{region 'Documentation'}
(*!
<summary>Reads a captured finding; the caller bounds the index by 8 subjects.</summary>
*)
{endregion}
METHOD PRIVATE IsFindingValid : BOOL //! TRUE when the selected captured finding satisfies the scenario metadata and diagnostic checks.
VAR_INPUT
    Index : UINT; //! One-based index in the retained isolated event capture.
    ExpectedName : STRING(GVL_Constants.NameLength); //! Independently authored Assertion name expected in the selected finding.
    ExpectedResult : E_Result; //! Independently authored finding result.
END_VAR
IsFindingValid := (FEvents[Index].SequenceId = UINT_TO_UDINT(Index))
    AND (FEvents[Index].Name = ExpectedName)
    AND (FEvents[Index].OwnerScope = E_OwnerScope.Assertion)
    AND (FEvents[Index].EventType = E_EventType.Result)
    AND (FEvents[Index].State = E_State.Running)
    AND (FEvents[Index].Result = ExpectedResult)
    AND (FEvents[Index].Message <> '');
END_METHOD

{region 'Documentation'}
(*!
<summary>Completes abort without asynchronous resources.</summary>
*)
{endregion}
METHOD PROTECTED ProcessAbort
VAR_INPUT
    Enable : BOOL; //! Phase permission supplied by the owning Test Case; FALSE does not authorize progression, while observation may continue.
END_VAR
IF Enable THEN
    CompleteAbort();
END_IF;
END_METHOD

{region 'Documentation'}
(*!
<summary>Latches checked observations before the next script step may proceed.</summary>
*)
{endregion}
METHOD PROTECTED ProcessAssertions
VAR_INPUT
    Enable : BOOL; //! Phase permission supplied by the owning Test Case; FALSE does not authorize progression, while observation may continue.
END_VAR
VAR
    Evaluate : BOOL;
END_VAR
Evaluate := Enable AND FObservationReady;
FEqualResult(Enable := Evaluate,
    State := State,
    IN := FEqualResultMatches);
FNotEqualResult(Enable := Evaluate,
    State := State,
    IN := FNotEqualResultMatches);
FLessThanResult(Enable := Evaluate,
    State := State,
    IN := FLessThanResultMatches);
FLessEqualResult(Enable := Evaluate,
    State := State,
    IN := FLessEqualResultMatches);
FGreaterThanResult(Enable := Evaluate,
    State := State,
    IN := FGreaterThanResultMatches);
FGreaterEqualResult(Enable := Evaluate,
    State := State,
    IN := FGreaterEqualResultMatches);
FInRangeResult(Enable := Evaluate,
    State := State,
    IN := FInRangeResultMatches);
FNotInRangeResult(Enable := Evaluate,
    State := State,
    IN := FNotInRangeResultMatches);
FCaptureIntegrity(Enable := Evaluate,
    State := State,
    IN := FCaptureIntegrityMatches);
FFindingDetails(Enable := Evaluate,
    State := State,
    IN := FFindingDetailsMatch);
IF Evaluate THEN
    FChecked := TRUE;
END_IF;
END_METHOD

{region 'Documentation'}
(*!
<summary>No Preparation phase is required.</summary>
*)
{endregion}
METHOD PROTECTED ProcessPreparations
VAR_INPUT
    // SA0033: Required hook; this test has no Preparation phase.
    {attribute 'analysis' := '-33'}
    Enable : BOOL; //! Phase permission supplied by the owning Test Case; FALSE does not authorize progression, while observation may continue.
END_VAR
END_METHOD

{region 'Documentation'}
(*!
<summary>Restarts the script and resets the checking Assertions.</summary>
*)
{endregion}
METHOD PROTECTED ProcessReset
FRow := EqualAtLowerBound;
FRowPrepared := FALSE;
FChecked := FALSE;
FObservationReady := FALSE;
FEqualResult.Reset();
FEqualResultMatches := TRUE;
FNotEqualResult.Reset();
FNotEqualResultMatches := TRUE;
FLessThanResult.Reset();
FLessThanResultMatches := TRUE;
FLessEqualResult.Reset();
FLessEqualResultMatches := TRUE;
FGreaterThanResult.Reset();
FGreaterThanResultMatches := TRUE;
FGreaterEqualResult.Reset();
FGreaterEqualResultMatches := TRUE;
FInRangeResult.Reset();
FInRangeResultMatches := TRUE;
FNotInRangeResult.Reset();
FNotInRangeResultMatches := TRUE;
FCaptureIntegrity.Reset();
FCaptureIntegrityMatches := TRUE;
FFindingDetails.Reset();
FFindingDetailsMatch := TRUE;
CompleteReset();
END_METHOD

{region 'Documentation'}
(*!
<summary>Advances one bounded script step per active PLC cycle.</summary>
*)
{endregion}
METHOD PROTECTED ProcessTests
VAR_INPUT
    Enable : BOOL; //! Phase permission supplied by the owning Test Case; FALSE does not authorize progression, while observation may continue.
END_VAR
IF NOT Enable THEN
    RETURN;
END_IF;

IF FChecked THEN
    FChecked := FALSE;
    FObservationReady := FALSE;
    IF FRow = LastRow THEN
        CompleteTests();
        RETURN;
    END_IF;
    FRow := FRow + 1;
    FRowPrepared := FALSE;
END_IF;

IF NOT FRowPrepared THEN
    SelectRow();
    FCapture.Reset();
    IF NOT FPreserveResults THEN
        ResetSubjects();
    END_IF;
    CallSubjects(Enable := FALSE);
    FRowPrepared := TRUE;
ELSE
    CallSubjects(Enable := TRUE);
    CheckResults();
    FObservationReady := TRUE;
END_IF;
END_METHOD

{region 'Documentation'}
(*!
<summary>Requests fresh subject results before the next disabled call.</summary>
*)
{endregion}
METHOD PRIVATE ResetSubjects
FEqualSubject.Reset();
FNotEqualSubject.Reset();
FLessThanSubject.Reset();
FLessEqualSubject.Reset();
FGreaterThanSubject.Reset();
FGreaterEqualSubject.Reset();
FInRangeSubject.Reset();
FNotInRangeSubject.Reset();
END_METHOD

{region 'Documentation'}
(*!
<summary>Selects independent literal outcomes; only named escalation rows preserve results.</summary>
*)
{endregion}
METHOD PRIVATE SelectRow
FPreserveResults := FALSE;
CASE FRow OF
    EqualAtLowerBound:
        FActual := REAL#1.0;
        FExpected := REAL#1.0;
        FLower := REAL#1.0;
        FUpper := REAL#2.0;
        FExpectedEqualResult := E_Result.Passed;
        FExpectedNotEqualResult := E_Result.Failed;
        FExpectedLessThanResult := E_Result.Failed;
        FExpectedLessEqualResult := E_Result.Passed;
        FExpectedGreaterThanResult := E_Result.Failed;
        FExpectedGreaterEqualResult := E_Result.Passed;
        FExpectedInRangeResult := E_Result.Passed;
        FExpectedNotInRangeResult := E_Result.Failed;
        FExpectedFindings := 4;
    AdjacentBelowExpected:
        FActual := REAL#1.0;
        FExpected := FAdjacent.Value;
        FLower := REAL#1.0;
        FUpper := FAdjacent.Value;
        FExpectedEqualResult := E_Result.Failed;
        FExpectedNotEqualResult := E_Result.Passed;
        FExpectedLessThanResult := E_Result.Passed;
        FExpectedLessEqualResult := E_Result.Passed;
        FExpectedGreaterThanResult := E_Result.Failed;
        FExpectedGreaterEqualResult := E_Result.Failed;
        FExpectedInRangeResult := E_Result.Passed;
        FExpectedNotInRangeResult := E_Result.Failed;
        FExpectedFindings := 4;
    AdjacentAboveExpected:
        FActual := FAdjacent.Value;
        FExpected := REAL#1.0;
        FLower := REAL#1.0;
        FUpper := FAdjacent.Value;
        FExpectedEqualResult := E_Result.Failed;
        FExpectedNotEqualResult := E_Result.Passed;
        FExpectedLessThanResult := E_Result.Failed;
        FExpectedLessEqualResult := E_Result.Failed;
        FExpectedGreaterThanResult := E_Result.Passed;
        FExpectedGreaterEqualResult := E_Result.Passed;
        FExpectedInRangeResult := E_Result.Passed;
        FExpectedNotInRangeResult := E_Result.Failed;
        FExpectedFindings := 4;
    Interior:
        FActual := REAL#1.5;
        FExpected := REAL#1.0;
        FLower := REAL#1.0;
        FUpper := REAL#2.0;
        FExpectedEqualResult := E_Result.Failed;
        FExpectedNotEqualResult := E_Result.Passed;
        FExpectedLessThanResult := E_Result.Failed;
        FExpectedLessEqualResult := E_Result.Failed;
        FExpectedGreaterThanResult := E_Result.Passed;
        FExpectedGreaterEqualResult := E_Result.Passed;
        FExpectedInRangeResult := E_Result.Passed;
        FExpectedNotInRangeResult := E_Result.Failed;
        FExpectedFindings := 4;
    BelowRange:
        FActual := REAL#0.0;
        FExpected := REAL#1.0;
        FLower := REAL#1.0;
        FUpper := REAL#2.0;
        FExpectedEqualResult := E_Result.Failed;
        FExpectedNotEqualResult := E_Result.Passed;
        FExpectedLessThanResult := E_Result.Passed;
        FExpectedLessEqualResult := E_Result.Passed;
        FExpectedGreaterThanResult := E_Result.Failed;
        FExpectedGreaterEqualResult := E_Result.Failed;
        FExpectedInRangeResult := E_Result.Failed;
        FExpectedNotInRangeResult := E_Result.Passed;
        FExpectedFindings := 4;
    AboveRange:
        FActual := REAL#3.0;
        FExpected := REAL#1.0;
        FLower := REAL#1.0;
        FUpper := REAL#2.0;
        FExpectedEqualResult := E_Result.Failed;
        FExpectedNotEqualResult := E_Result.Passed;
        FExpectedLessThanResult := E_Result.Failed;
        FExpectedLessEqualResult := E_Result.Failed;
        FExpectedGreaterThanResult := E_Result.Passed;
        FExpectedGreaterEqualResult := E_Result.Passed;
        FExpectedInRangeResult := E_Result.Failed;
        FExpectedNotInRangeResult := E_Result.Passed;
        FExpectedFindings := 4;
    EqualBounds:
        FActual := REAL#1.0;
        FExpected := REAL#1.0;
        FLower := REAL#1.0;
        FUpper := REAL#1.0;
        FExpectedEqualResult := E_Result.Passed;
        FExpectedNotEqualResult := E_Result.Failed;
        FExpectedLessThanResult := E_Result.Failed;
        FExpectedLessEqualResult := E_Result.Passed;
        FExpectedGreaterThanResult := E_Result.Failed;
        FExpectedGreaterEqualResult := E_Result.Passed;
        FExpectedInRangeResult := E_Result.Passed;
        FExpectedNotInRangeResult := E_Result.Failed;
        FExpectedFindings := 4;
    ReversedBounds:
        FActual := REAL#1.0;
        FExpected := REAL#1.0;
        FLower := REAL#2.0;
        FUpper := REAL#1.0;
        FExpectedEqualResult := E_Result.Passed;
        FExpectedNotEqualResult := E_Result.Failed;
        FExpectedLessThanResult := E_Result.Failed;
        FExpectedLessEqualResult := E_Result.Passed;
        FExpectedGreaterThanResult := E_Result.Failed;
        FExpectedGreaterEqualResult := E_Result.Passed;
        FExpectedInRangeResult := E_Result.Error;
        FExpectedNotInRangeResult := E_Result.Error;
        FExpectedFindings := 5;
    SignedZero:
        FActual := FNegativeZero.Value;
        FExpected := REAL#0.0;
        FLower := REAL#0.0;
        FUpper := REAL#0.0;
        FExpectedEqualResult := E_Result.Passed;
        FExpectedNotEqualResult := E_Result.Failed;
        FExpectedLessThanResult := E_Result.Failed;
        FExpectedLessEqualResult := E_Result.Passed;
        FExpectedGreaterThanResult := E_Result.Failed;
        FExpectedGreaterEqualResult := E_Result.Passed;
        FExpectedInRangeResult := E_Result.Passed;
        FExpectedNotInRangeResult := E_Result.Failed;
        FExpectedFindings := 4;
    ExtremeAscending:
        FActual := -FMaximum.Value;
        FExpected := FMaximum.Value;
        FLower := -FMaximum.Value;
        FUpper := FMaximum.Value;
        FExpectedEqualResult := E_Result.Failed;
        FExpectedNotEqualResult := E_Result.Passed;
        FExpectedLessThanResult := E_Result.Passed;
        FExpectedLessEqualResult := E_Result.Passed;
        FExpectedGreaterThanResult := E_Result.Failed;
        FExpectedGreaterEqualResult := E_Result.Failed;
        FExpectedInRangeResult := E_Result.Passed;
        FExpectedNotInRangeResult := E_Result.Failed;
        FExpectedFindings := 4;
    ExtremeDescending:
        FActual := FMaximum.Value;
        FExpected := -FMaximum.Value;
        FLower := -FMaximum.Value;
        FUpper := FMaximum.Value;
        FExpectedEqualResult := E_Result.Failed;
        FExpectedNotEqualResult := E_Result.Passed;
        FExpectedLessThanResult := E_Result.Failed;
        FExpectedLessEqualResult := E_Result.Failed;
        FExpectedGreaterThanResult := E_Result.Passed;
        FExpectedGreaterEqualResult := E_Result.Passed;
        FExpectedInRangeResult := E_Result.Passed;
        FExpectedNotInRangeResult := E_Result.Failed;
        FExpectedFindings := 4;
ELSE
    Error(Message := 'Unknown floating-point test row.');
END_CASE;
END_METHOD

END_FUNCTION_BLOCK

// ---- SelfTests/TestCases/TestSuite_AssertionFloatingPoint/Test_AssertionRelations_LReal.TcPOU
{region 'Documentation'}
(*!
<summary>Checks exact LREAL ordering, inclusive ranges and signed zero.</summary>
<description>
Adjacent values differ by one representable step above 1; no implicit epsilon is allowed.
Range rows include both endpoints, equal bounds and invalid reversed bounds.
Extreme ordering uses comparisons only, not arithmetic differences.
A disabled preparation call consumes subject resets before the next enabled observation.
Only outer checking Assertions contribute to the Test Case result.
Expected outcomes are explicit; production processing is inherited, not mirrored.
</description>
*)
{endregion}
FUNCTION_BLOCK Test_AssertionRelations_LReal EXTENDS TestCaseBase
VAR
    FEqualSubject : AssertEqual_LReal;
    FNotEqualSubject : AssertNotEqual_LReal;
    FLessThanSubject : AssertLessThan_LReal;
    FLessEqualSubject : AssertLessEqual_LReal;
    FGreaterThanSubject : AssertGreaterThan_LReal;
    FGreaterEqualSubject : AssertGreaterEqual_LReal;
    FInRangeSubject : AssertInRange_LReal;
    FNotInRangeSubject : AssertNotInRange_LReal;
    FActual : LREAL;
    FExpected : LREAL;
    FLower : LREAL;
    FUpper : LREAL;
    FMaximum : FloatingPointBits_LReal;
    FAdjacent : FloatingPointBits_LReal;
    FNegativeZero : FloatingPointBits_LReal;
    FExpectedEqualResult : E_Result;
    FExpectedNotEqualResult : E_Result;
    FExpectedLessThanResult : E_Result;
    FExpectedLessEqualResult : E_Result;
    FExpectedGreaterThanResult : E_Result;
    FExpectedGreaterEqualResult : E_Result;
    FExpectedInRangeResult : E_Result;
    FExpectedNotInRangeResult : E_Result;
    FExpectedFindings : UDINT;
    FCapture : EventBuffer;
    FEvents : ARRAY[1..CaptureLength] OF ST_Event;
    FCaptureFifo : ST_FifoStatus;
    FCaptureStatus : ST_EventBufferStatus;
    FRow : UINT;
    FRowPrepared : BOOL;
    FPreserveResults : BOOL;
    FObservationReady : BOOL;
    FChecked : BOOL;
    FSetupValid : BOOL;
END_VAR
VAR
    FEqualResult : AssertTrue;
    FEqualResultMatches : BOOL;
    FNotEqualResult : AssertTrue;
    FNotEqualResultMatches : BOOL;
    FLessThanResult : AssertTrue;
    FLessThanResultMatches : BOOL;
    FLessEqualResult : AssertTrue;
    FLessEqualResultMatches : BOOL;
    FGreaterThanResult : AssertTrue;
    FGreaterThanResultMatches : BOOL;
    FGreaterEqualResult : AssertTrue;
    FGreaterEqualResultMatches : BOOL;
    FInRangeResult : AssertTrue;
    FInRangeResultMatches : BOOL;
    FNotInRangeResult : AssertTrue;
    FNotInRangeResultMatches : BOOL;
    FCaptureIntegrity : AssertTrue;
    FCaptureIntegrityMatches : BOOL;
    FFindingDetails : AssertTrue;
    FFindingDetailsMatch : BOOL;
END_VAR
VAR CONSTANT
    CaptureLength : UINT := 16;
    FixtureSize : UINT := 8;
    OneBits : LWORD := LWORD#16#3FF0000000000000;
    MaximumBits : LWORD := LWORD#16#7FEFFFFFFFFFFFFF;
    AdjacentBits : LWORD := LWORD#16#3FF0000000000001;
    NegativeZeroBits : LWORD := LWORD#16#8000000000000000;
    EqualAtLowerBound : UINT := 1;
    AdjacentBelowExpected : UINT := 2;
    AdjacentAboveExpected : UINT := 3;
    Interior : UINT := 4;
    BelowRange : UINT := 5;
    AboveRange : UINT := 6;
    EqualBounds : UINT := 7;
    ReversedBounds : UINT := 8;
    SignedZero : UINT := 9;
    ExtremeAscending : UINT := 10;
    ExtremeDescending : UINT := 11;
    LastRow : UINT := ExtremeDescending;
END_VAR

SUPER^();

{region 'Documentation'}
(*!
<summary>Collects only outer checking Assertions, never intentional subject findings.</summary>
*)
{endregion}
METHOD PROTECTED AggregateResults
VAR_INPUT
    Aggregator : I_ResultAggregator; //! Borrowed result sink owned by the outer Test Case; add this test's checking Assertions without resetting or retaining the sink.
END_VAR
Aggregator.AddProvider(Provider := FEqualResult);
Aggregator.AddProvider(Provider := FNotEqualResult);
Aggregator.AddProvider(Provider := FLessThanResult);
Aggregator.AddProvider(Provider := FLessEqualResult);
Aggregator.AddProvider(Provider := FGreaterThanResult);
Aggregator.AddProvider(Provider := FGreaterEqualResult);
Aggregator.AddProvider(Provider := FInRangeResult);
Aggregator.AddProvider(Provider := FNotInRangeResult);
Aggregator.AddProvider(Provider := FCaptureIntegrity);
Aggregator.AddProvider(Provider := FFindingDetails);
END_METHOD

{region 'Documentation'}
(*!
<summary>Calls each inherited production Assertion once using the selected row.</summary>
*)
{endregion}
METHOD PRIVATE CallSubjects
VAR_INPUT
    Enable : BOOL; //! Observation-enable input forwarded to the controlled Assertion subjects for this call.
END_VAR
FEqualSubject(Enable := Enable,
    State := E_State.Running,
    IN := FActual,
    Expected := FExpected);
FNotEqualSubject(Enable := Enable,
    State := E_State.Running,
    IN := FActual,
    Expected := FExpected);
FLessThanSubject(Enable := Enable,
    State := E_State.Running,
    IN := FActual,
    Maximum := FExpected);
FLessEqualSubject(Enable := Enable,
    State := E_State.Running,
    IN := FActual,
    Maximum := FExpected);
FGreaterThanSubject(Enable := Enable,
    State := E_State.Running,
    IN := FActual,
    Minimum := FExpected);
FGreaterEqualSubject(Enable := Enable,
    State := E_State.Running,
    IN := FActual,
    Minimum := FExpected);
FInRangeSubject(Enable := Enable,
    State := E_State.Running,
    IN := FActual,
    Minimum := FLower,
    Maximum := FUpper);
FNotInRangeSubject(Enable := Enable,
    State := E_State.Running,
    IN := FActual,
    Minimum := FLower,
    Maximum := FUpper);
END_METHOD

{region 'Documentation'}
(*!
<summary>Extends base validation with subject and checking-Assertion setup.</summary>
*)
{endregion}
METHOD PROTECTED CheckInitialization : BOOL //! TRUE when the inherited initialization check and this concrete fixture check both accept the setup.
CheckInitialization := SUPER^.CheckInitialization();
IF NOT CheckInitialization THEN
    RETURN;
END_IF;

CheckInitialization := FSetupValid
    AND FEqualResult.IsInitialized
    AND FNotEqualResult.IsInitialized
    AND FLessThanResult.IsInitialized
    AND FLessEqualResult.IsInitialized
    AND FGreaterThanResult.IsInitialized
    AND FGreaterEqualResult.IsInitialized
    AND FInRangeResult.IsInitialized
    AND FNotInRangeResult.IsInitialized
    AND FCaptureIntegrity.IsInitialized
    AND FFindingDetails.IsInitialized;
IF NOT CheckInitialization THEN
    EventPublisher.PublishEvent(Event := CreateFrameworkEvent(Name := Name,
        ResourceName := '',
        State := State,
        Severity := E_EventSeverity.Error,
        Message := 'Floating-point selftest setup or fixture representation failed.'));
END_IF;
END_METHOD

{region 'Documentation'}
(*!
<summary>Checks literal results and the ordered isolated findings from this row.</summary>
*)
{endregion}
METHOD PRIVATE CheckResults
VAR
    FindingIndex : UINT;
    FindingMatches : BOOL;
END_VAR
FEqualResultMatches := FEqualSubject.Result = FExpectedEqualResult;
FNotEqualResultMatches := FNotEqualSubject.Result = FExpectedNotEqualResult;
FLessThanResultMatches := FLessThanSubject.Result = FExpectedLessThanResult;
FLessEqualResultMatches := FLessEqualSubject.Result = FExpectedLessEqualResult;
FGreaterThanResultMatches := FGreaterThanSubject.Result = FExpectedGreaterThanResult;
FGreaterEqualResultMatches := FGreaterEqualSubject.Result = FExpectedGreaterEqualResult;
FInRangeResultMatches := FInRangeSubject.Result = FExpectedInRangeResult;
FNotInRangeResultMatches := FNotInRangeSubject.Result = FExpectedNotInRangeResult;
FCaptureIntegrityMatches := (FCaptureStatus.SequenceId = FExpectedFindings)
    AND (FCaptureStatus.LostEventCount = 0);

FindingIndex := 1;
FFindingDetailsMatch := TRUE;
IF (FExpectedEqualResult = E_Result.Failed) OR (FExpectedEqualResult = E_Result.Error) THEN
    FindingMatches := IsFindingValid(Index := FindingIndex,
        ExpectedName := FEqualSubject.Name,
        ExpectedResult := FExpectedEqualResult);
    FFindingDetailsMatch := FFindingDetailsMatch AND FindingMatches;
    FindingIndex := FindingIndex + 1;
END_IF;
IF (FExpectedNotEqualResult = E_Result.Failed) OR (FExpectedNotEqualResult = E_Result.Error) THEN
    FindingMatches := IsFindingValid(Index := FindingIndex,
        ExpectedName := FNotEqualSubject.Name,
        ExpectedResult := FExpectedNotEqualResult);
    FFindingDetailsMatch := FFindingDetailsMatch AND FindingMatches;
    FindingIndex := FindingIndex + 1;
END_IF;
IF (FExpectedLessThanResult = E_Result.Failed) OR (FExpectedLessThanResult = E_Result.Error) THEN
    FindingMatches := IsFindingValid(Index := FindingIndex,
        ExpectedName := FLessThanSubject.Name,
        ExpectedResult := FExpectedLessThanResult);
    FFindingDetailsMatch := FFindingDetailsMatch AND FindingMatches;
    FindingIndex := FindingIndex + 1;
END_IF;
IF (FExpectedLessEqualResult = E_Result.Failed) OR (FExpectedLessEqualResult = E_Result.Error) THEN
    FindingMatches := IsFindingValid(Index := FindingIndex,
        ExpectedName := FLessEqualSubject.Name,
        ExpectedResult := FExpectedLessEqualResult);
    FFindingDetailsMatch := FFindingDetailsMatch AND FindingMatches;
    FindingIndex := FindingIndex + 1;
END_IF;
IF (FExpectedGreaterThanResult = E_Result.Failed) OR (FExpectedGreaterThanResult = E_Result.Error) THEN
    FindingMatches := IsFindingValid(Index := FindingIndex,
        ExpectedName := FGreaterThanSubject.Name,
        ExpectedResult := FExpectedGreaterThanResult);
    FFindingDetailsMatch := FFindingDetailsMatch AND FindingMatches;
    FindingIndex := FindingIndex + 1;
END_IF;
IF (FExpectedGreaterEqualResult = E_Result.Failed) OR (FExpectedGreaterEqualResult = E_Result.Error) THEN
    FindingMatches := IsFindingValid(Index := FindingIndex,
        ExpectedName := FGreaterEqualSubject.Name,
        ExpectedResult := FExpectedGreaterEqualResult);
    FFindingDetailsMatch := FFindingDetailsMatch AND FindingMatches;
    FindingIndex := FindingIndex + 1;
END_IF;
IF (FExpectedInRangeResult = E_Result.Failed) OR (FExpectedInRangeResult = E_Result.Error) THEN
    FindingMatches := IsFindingValid(Index := FindingIndex,
        ExpectedName := FInRangeSubject.Name,
        ExpectedResult := FExpectedInRangeResult);
    FFindingDetailsMatch := FFindingDetailsMatch AND FindingMatches;
    FindingIndex := FindingIndex + 1;
END_IF;
IF (FExpectedNotInRangeResult = E_Result.Failed) OR (FExpectedNotInRangeResult = E_Result.Error) THEN
    FindingMatches := IsFindingValid(Index := FindingIndex,
        ExpectedName := FNotInRangeSubject.Name,
        ExpectedResult := FExpectedNotInRangeResult);
    FFindingDetailsMatch := FFindingDetailsMatch AND FindingMatches;
    FindingIndex := FindingIndex + 1;
END_IF;
END_METHOD

{region 'Documentation'}
(*!
<summary>Configures checking Assertions; subject actions remain in the test script.</summary>
*)
{endregion}
METHOD PROTECTED Configure
VAR
    Initialized : BOOL;
END_VAR
FPreparationStateCount := 0;
FTestStateCount := 1;
FSetupValid := InitializeValues();
FEqualResult.Initialize(Parent := THIS^,
    AssertionName := 'EqualResult');
FNotEqualResult.Initialize(Parent := THIS^,
    AssertionName := 'NotEqualResult');
FLessThanResult.Initialize(Parent := THIS^,
    AssertionName := 'LessThanResult');
FLessEqualResult.Initialize(Parent := THIS^,
    AssertionName := 'LessEqualResult');
FGreaterThanResult.Initialize(Parent := THIS^,
    AssertionName := 'GreaterThanResult');
FGreaterEqualResult.Initialize(Parent := THIS^,
    AssertionName := 'GreaterEqualResult');
FInRangeResult.Initialize(Parent := THIS^,
    AssertionName := 'InRangeResult');
FNotInRangeResult.Initialize(Parent := THIS^,
    AssertionName := 'NotInRangeResult');
FCaptureIntegrity.Initialize(Parent := THIS^,
    AssertionName := 'CaptureIntegrity');
FFindingDetails.Initialize(Parent := THIS^,
    AssertionName := 'FindingDetails');
Initialized := FCapture.Initialize(Buffer := FEvents,
    FifoControl := FCaptureFifo,
    Status := FCaptureStatus);
FSetupValid := FSetupValid AND Initialized;
FEqualSubject.BindPublisher(Publisher := FCapture);
Initialized := FEqualSubject.Initialize(Parent := THIS^,
    AssertionName := 'EqualSubject');
FSetupValid := FSetupValid AND Initialized;
FNotEqualSubject.BindPublisher(Publisher := FCapture);
Initialized := FNotEqualSubject.Initialize(Parent := THIS^,
    AssertionName := 'NotEqualSubject');
FSetupValid := FSetupValid AND Initialized;
FLessThanSubject.BindPublisher(Publisher := FCapture);
Initialized := FLessThanSubject.Initialize(Parent := THIS^,
    AssertionName := 'LessThanSubject');
FSetupValid := FSetupValid AND Initialized;
FLessEqualSubject.BindPublisher(Publisher := FCapture);
Initialized := FLessEqualSubject.Initialize(Parent := THIS^,
    AssertionName := 'LessEqualSubject');
FSetupValid := FSetupValid AND Initialized;
FGreaterThanSubject.BindPublisher(Publisher := FCapture);
Initialized := FGreaterThanSubject.Initialize(Parent := THIS^,
    AssertionName := 'GreaterThanSubject');
FSetupValid := FSetupValid AND Initialized;
FGreaterEqualSubject.BindPublisher(Publisher := FCapture);
Initialized := FGreaterEqualSubject.Initialize(Parent := THIS^,
    AssertionName := 'GreaterEqualSubject');
FSetupValid := FSetupValid AND Initialized;
FInRangeSubject.BindPublisher(Publisher := FCapture);
Initialized := FInRangeSubject.Initialize(Parent := THIS^,
    AssertionName := 'InRangeSubject');
FSetupValid := FSetupValid AND Initialized;
FNotInRangeSubject.BindPublisher(Publisher := FCapture);
Initialized := FNotInRangeSubject.Initialize(Parent := THIS^,
    AssertionName := 'NotInRangeSubject');
FSetupValid := FSetupValid AND Initialized;
END_METHOD

{region 'Documentation'}
(*!
<summary>Establishes typed fixtures and verifies their representation before any subject call.</summary>
*)
{endregion}
METHOD PRIVATE InitializeValues : BOOL //! TRUE when fixture sizes and floating-point bit representations match their explicit expected patterns.
VAR
    Representation : FloatingPointBits_LReal;
END_VAR
Representation.Value := LREAL#1.0;
InitializeValues := (SIZEOF(Representation) = FixtureSize)
    AND (Representation.Bits = OneBits);

FMaximum.Value := LREAL#1.7976931348623157E308;
Representation.Value := FMaximum.Value;
InitializeValues := InitializeValues AND (Representation.Bits = MaximumBits);
FAdjacent.Value := LREAL#1.0000000000000002220446049250313080847263336181640625;
Representation.Value := FAdjacent.Value;
InitializeValues := InitializeValues AND (Representation.Bits = AdjacentBits);
FNegativeZero.Bits := NegativeZeroBits;
Representation.Value := FNegativeZero.Value;
InitializeValues := InitializeValues AND (Representation.Bits = NegativeZeroBits);
END_METHOD

{region 'Documentation'}
(*!
<summary>Reads a captured finding; the caller bounds the index by 8 subjects.</summary>
*)
{endregion}
METHOD PRIVATE IsFindingValid : BOOL //! TRUE when the selected captured finding satisfies the scenario metadata and diagnostic checks.
VAR_INPUT
    Index : UINT; //! One-based index in the retained isolated event capture.
    ExpectedName : STRING(GVL_Constants.NameLength); //! Independently authored Assertion name expected in the selected finding.
    ExpectedResult : E_Result; //! Independently authored finding result.
END_VAR
IsFindingValid := (FEvents[Index].SequenceId = UINT_TO_UDINT(Index))
    AND (FEvents[Index].Name = ExpectedName)
    AND (FEvents[Index].OwnerScope = E_OwnerScope.Assertion)
    AND (FEvents[Index].EventType = E_EventType.Result)
    AND (FEvents[Index].State = E_State.Running)
    AND (FEvents[Index].Result = ExpectedResult)
    AND (FEvents[Index].Message <> '');
END_METHOD

{region 'Documentation'}
(*!
<summary>Completes abort without asynchronous resources.</summary>
*)
{endregion}
METHOD PROTECTED ProcessAbort
VAR_INPUT
    Enable : BOOL; //! Phase permission supplied by the owning Test Case; FALSE does not authorize progression, while observation may continue.
END_VAR
IF Enable THEN
    CompleteAbort();
END_IF;
END_METHOD

{region 'Documentation'}
(*!
<summary>Latches checked observations before the next script step may proceed.</summary>
*)
{endregion}
METHOD PROTECTED ProcessAssertions
VAR_INPUT
    Enable : BOOL; //! Phase permission supplied by the owning Test Case; FALSE does not authorize progression, while observation may continue.
END_VAR
VAR
    Evaluate : BOOL;
END_VAR
Evaluate := Enable AND FObservationReady;
FEqualResult(Enable := Evaluate,
    State := State,
    IN := FEqualResultMatches);
FNotEqualResult(Enable := Evaluate,
    State := State,
    IN := FNotEqualResultMatches);
FLessThanResult(Enable := Evaluate,
    State := State,
    IN := FLessThanResultMatches);
FLessEqualResult(Enable := Evaluate,
    State := State,
    IN := FLessEqualResultMatches);
FGreaterThanResult(Enable := Evaluate,
    State := State,
    IN := FGreaterThanResultMatches);
FGreaterEqualResult(Enable := Evaluate,
    State := State,
    IN := FGreaterEqualResultMatches);
FInRangeResult(Enable := Evaluate,
    State := State,
    IN := FInRangeResultMatches);
FNotInRangeResult(Enable := Evaluate,
    State := State,
    IN := FNotInRangeResultMatches);
FCaptureIntegrity(Enable := Evaluate,
    State := State,
    IN := FCaptureIntegrityMatches);
FFindingDetails(Enable := Evaluate,
    State := State,
    IN := FFindingDetailsMatch);
IF Evaluate THEN
    FChecked := TRUE;
END_IF;
END_METHOD

{region 'Documentation'}
(*!
<summary>No Preparation phase is required.</summary>
*)
{endregion}
METHOD PROTECTED ProcessPreparations
VAR_INPUT
    // SA0033: Required hook; this test has no Preparation phase.
    {attribute 'analysis' := '-33'}
    Enable : BOOL; //! Phase permission supplied by the owning Test Case; FALSE does not authorize progression, while observation may continue.
END_VAR
END_METHOD

{region 'Documentation'}
(*!
<summary>Restarts the script and resets the checking Assertions.</summary>
*)
{endregion}
METHOD PROTECTED ProcessReset
FRow := EqualAtLowerBound;
FRowPrepared := FALSE;
FChecked := FALSE;
FObservationReady := FALSE;
FEqualResult.Reset();
FEqualResultMatches := TRUE;
FNotEqualResult.Reset();
FNotEqualResultMatches := TRUE;
FLessThanResult.Reset();
FLessThanResultMatches := TRUE;
FLessEqualResult.Reset();
FLessEqualResultMatches := TRUE;
FGreaterThanResult.Reset();
FGreaterThanResultMatches := TRUE;
FGreaterEqualResult.Reset();
FGreaterEqualResultMatches := TRUE;
FInRangeResult.Reset();
FInRangeResultMatches := TRUE;
FNotInRangeResult.Reset();
FNotInRangeResultMatches := TRUE;
FCaptureIntegrity.Reset();
FCaptureIntegrityMatches := TRUE;
FFindingDetails.Reset();
FFindingDetailsMatch := TRUE;
CompleteReset();
END_METHOD

{region 'Documentation'}
(*!
<summary>Advances one bounded script step per active PLC cycle.</summary>
*)
{endregion}
METHOD PROTECTED ProcessTests
VAR_INPUT
    Enable : BOOL; //! Phase permission supplied by the owning Test Case; FALSE does not authorize progression, while observation may continue.
END_VAR
IF NOT Enable THEN
    RETURN;
END_IF;

IF FChecked THEN
    FChecked := FALSE;
    FObservationReady := FALSE;
    IF FRow = LastRow THEN
        CompleteTests();
        RETURN;
    END_IF;
    FRow := FRow + 1;
    FRowPrepared := FALSE;
END_IF;

IF NOT FRowPrepared THEN
    SelectRow();
    FCapture.Reset();
    IF NOT FPreserveResults THEN
        ResetSubjects();
    END_IF;
    CallSubjects(Enable := FALSE);
    FRowPrepared := TRUE;
ELSE
    CallSubjects(Enable := TRUE);
    CheckResults();
    FObservationReady := TRUE;
END_IF;
END_METHOD

{region 'Documentation'}
(*!
<summary>Requests fresh subject results before the next disabled call.</summary>
*)
{endregion}
METHOD PRIVATE ResetSubjects
FEqualSubject.Reset();
FNotEqualSubject.Reset();
FLessThanSubject.Reset();
FLessEqualSubject.Reset();
FGreaterThanSubject.Reset();
FGreaterEqualSubject.Reset();
FInRangeSubject.Reset();
FNotInRangeSubject.Reset();
END_METHOD

{region 'Documentation'}
(*!
<summary>Selects independent literal outcomes; only named escalation rows preserve results.</summary>
*)
{endregion}
METHOD PRIVATE SelectRow
FPreserveResults := FALSE;
CASE FRow OF
    EqualAtLowerBound:
        FActual := LREAL#1.0;
        FExpected := LREAL#1.0;
        FLower := LREAL#1.0;
        FUpper := LREAL#2.0;
        FExpectedEqualResult := E_Result.Passed;
        FExpectedNotEqualResult := E_Result.Failed;
        FExpectedLessThanResult := E_Result.Failed;
        FExpectedLessEqualResult := E_Result.Passed;
        FExpectedGreaterThanResult := E_Result.Failed;
        FExpectedGreaterEqualResult := E_Result.Passed;
        FExpectedInRangeResult := E_Result.Passed;
        FExpectedNotInRangeResult := E_Result.Failed;
        FExpectedFindings := 4;
    AdjacentBelowExpected:
        FActual := LREAL#1.0;
        FExpected := FAdjacent.Value;
        FLower := LREAL#1.0;
        FUpper := FAdjacent.Value;
        FExpectedEqualResult := E_Result.Failed;
        FExpectedNotEqualResult := E_Result.Passed;
        FExpectedLessThanResult := E_Result.Passed;
        FExpectedLessEqualResult := E_Result.Passed;
        FExpectedGreaterThanResult := E_Result.Failed;
        FExpectedGreaterEqualResult := E_Result.Failed;
        FExpectedInRangeResult := E_Result.Passed;
        FExpectedNotInRangeResult := E_Result.Failed;
        FExpectedFindings := 4;
    AdjacentAboveExpected:
        FActual := FAdjacent.Value;
        FExpected := LREAL#1.0;
        FLower := LREAL#1.0;
        FUpper := FAdjacent.Value;
        FExpectedEqualResult := E_Result.Failed;
        FExpectedNotEqualResult := E_Result.Passed;
        FExpectedLessThanResult := E_Result.Failed;
        FExpectedLessEqualResult := E_Result.Failed;
        FExpectedGreaterThanResult := E_Result.Passed;
        FExpectedGreaterEqualResult := E_Result.Passed;
        FExpectedInRangeResult := E_Result.Passed;
        FExpectedNotInRangeResult := E_Result.Failed;
        FExpectedFindings := 4;
    Interior:
        FActual := LREAL#1.5;
        FExpected := LREAL#1.0;
        FLower := LREAL#1.0;
        FUpper := LREAL#2.0;
        FExpectedEqualResult := E_Result.Failed;
        FExpectedNotEqualResult := E_Result.Passed;
        FExpectedLessThanResult := E_Result.Failed;
        FExpectedLessEqualResult := E_Result.Failed;
        FExpectedGreaterThanResult := E_Result.Passed;
        FExpectedGreaterEqualResult := E_Result.Passed;
        FExpectedInRangeResult := E_Result.Passed;
        FExpectedNotInRangeResult := E_Result.Failed;
        FExpectedFindings := 4;
    BelowRange:
        FActual := LREAL#0.0;
        FExpected := LREAL#1.0;
        FLower := LREAL#1.0;
        FUpper := LREAL#2.0;
        FExpectedEqualResult := E_Result.Failed;
        FExpectedNotEqualResult := E_Result.Passed;
        FExpectedLessThanResult := E_Result.Passed;
        FExpectedLessEqualResult := E_Result.Passed;
        FExpectedGreaterThanResult := E_Result.Failed;
        FExpectedGreaterEqualResult := E_Result.Failed;
        FExpectedInRangeResult := E_Result.Failed;
        FExpectedNotInRangeResult := E_Result.Passed;
        FExpectedFindings := 4;
    AboveRange:
        FActual := LREAL#3.0;
        FExpected := LREAL#1.0;
        FLower := LREAL#1.0;
        FUpper := LREAL#2.0;
        FExpectedEqualResult := E_Result.Failed;
        FExpectedNotEqualResult := E_Result.Passed;
        FExpectedLessThanResult := E_Result.Failed;
        FExpectedLessEqualResult := E_Result.Failed;
        FExpectedGreaterThanResult := E_Result.Passed;
        FExpectedGreaterEqualResult := E_Result.Passed;
        FExpectedInRangeResult := E_Result.Failed;
        FExpectedNotInRangeResult := E_Result.Passed;
        FExpectedFindings := 4;
    EqualBounds:
        FActual := LREAL#1.0;
        FExpected := LREAL#1.0;
        FLower := LREAL#1.0;
        FUpper := LREAL#1.0;
        FExpectedEqualResult := E_Result.Passed;
        FExpectedNotEqualResult := E_Result.Failed;
        FExpectedLessThanResult := E_Result.Failed;
        FExpectedLessEqualResult := E_Result.Passed;
        FExpectedGreaterThanResult := E_Result.Failed;
        FExpectedGreaterEqualResult := E_Result.Passed;
        FExpectedInRangeResult := E_Result.Passed;
        FExpectedNotInRangeResult := E_Result.Failed;
        FExpectedFindings := 4;
    ReversedBounds:
        FActual := LREAL#1.0;
        FExpected := LREAL#1.0;
        FLower := LREAL#2.0;
        FUpper := LREAL#1.0;
        FExpectedEqualResult := E_Result.Passed;
        FExpectedNotEqualResult := E_Result.Failed;
        FExpectedLessThanResult := E_Result.Failed;
        FExpectedLessEqualResult := E_Result.Passed;
        FExpectedGreaterThanResult := E_Result.Failed;
        FExpectedGreaterEqualResult := E_Result.Passed;
        FExpectedInRangeResult := E_Result.Error;
        FExpectedNotInRangeResult := E_Result.Error;
        FExpectedFindings := 5;
    SignedZero:
        FActual := FNegativeZero.Value;
        FExpected := LREAL#0.0;
        FLower := LREAL#0.0;
        FUpper := LREAL#0.0;
        FExpectedEqualResult := E_Result.Passed;
        FExpectedNotEqualResult := E_Result.Failed;
        FExpectedLessThanResult := E_Result.Failed;
        FExpectedLessEqualResult := E_Result.Passed;
        FExpectedGreaterThanResult := E_Result.Failed;
        FExpectedGreaterEqualResult := E_Result.Passed;
        FExpectedInRangeResult := E_Result.Passed;
        FExpectedNotInRangeResult := E_Result.Failed;
        FExpectedFindings := 4;
    ExtremeAscending:
        FActual := -FMaximum.Value;
        FExpected := FMaximum.Value;
        FLower := -FMaximum.Value;
        FUpper := FMaximum.Value;
        FExpectedEqualResult := E_Result.Failed;
        FExpectedNotEqualResult := E_Result.Passed;
        FExpectedLessThanResult := E_Result.Passed;
        FExpectedLessEqualResult := E_Result.Passed;
        FExpectedGreaterThanResult := E_Result.Failed;
        FExpectedGreaterEqualResult := E_Result.Failed;
        FExpectedInRangeResult := E_Result.Passed;
        FExpectedNotInRangeResult := E_Result.Failed;
        FExpectedFindings := 4;
    ExtremeDescending:
        FActual := FMaximum.Value;
        FExpected := -FMaximum.Value;
        FLower := -FMaximum.Value;
        FUpper := FMaximum.Value;
        FExpectedEqualResult := E_Result.Failed;
        FExpectedNotEqualResult := E_Result.Passed;
        FExpectedLessThanResult := E_Result.Failed;
        FExpectedLessEqualResult := E_Result.Failed;
        FExpectedGreaterThanResult := E_Result.Passed;
        FExpectedGreaterEqualResult := E_Result.Passed;
        FExpectedInRangeResult := E_Result.Passed;
        FExpectedNotInRangeResult := E_Result.Failed;
        FExpectedFindings := 4;
ELSE
    Error(Message := 'Unknown floating-point test row.');
END_CASE;
END_METHOD

END_FUNCTION_BLOCK

// ---- Framework/Assertions/POU/BasicTypes/LReal/AssertEqual_LReal.TcPOU
{region 'Documentation'}
(*!
<summary>Checks equality with the expected LREAL value.</summary>
<description>

All checked operands and bounds must be finite; NaN or either infinity reports Error
during active evaluation.

Numeric diagnostics use the formatter's default six significant digits; rounding affects
the message only, not the comparison.

</description>
*)
{endregion}
FUNCTION_BLOCK AssertEqual_LReal EXTENDS AssertionBase
VAR_INPUT
    IN : LREAL; //! Actual value checked or observed by this Assertion.
    Expected : LREAL; //! Reference value for comparison with IN.
END_VAR

SUPER^();

{region 'Documentation'}
(*!
<summary>Check equality with the expected LREAL value.</summary>
*)
{endregion}
METHOD PROTECTED Assert
VAR
    Message : STRING(GVL_Constants.MessageLength);
    ExpectedText : STRING(GVL_Constants.AssertionValueLength);
    ActualText : STRING(GVL_Constants.AssertionValueLength);
END_VAR
IF NOT EvaluationActive THEN
    RETURN;
END_IF;

IF Result = E_Result.Error THEN
    RETURN;
END_IF;

IF NOT Tc2_Utilities.LrealIsFinite(x := IN) THEN
    Error(Message := 'Assertion error: IN must be finite.');
    RETURN;
END_IF;

IF NOT Tc2_Utilities.LrealIsFinite(x := Expected) THEN
    Error(Message := 'Assertion error: Expected must be finite.');
    RETURN;
END_IF;

IF Result = E_Result.Failed THEN
    RETURN;
END_IF;

IF IN <> Expected THEN
    ExpectedText := CreateAssertionTextValue_LReal(Value := Expected);
    ActualText := CreateAssertionTextValue_LReal(Value := IN);
    Message := CONCAT('Assertion failed: values are not equal. Expected = ',
        ExpectedText);
    Message := CONCAT(Message, ', Actual = ');
    Message := CONCAT(Message, ActualText);
    Message := CONCAT(Message, '.');
    Fail(Message := Message);
    RETURN;
END_IF;

Pass();
END_METHOD

END_FUNCTION_BLOCK

// ---- Framework/Assertions/POU/BasicTypes/LReal/AssertNotEqual_LReal.TcPOU
{region 'Documentation'}
(*!
<summary>Checks inequality with the forbidden LREAL value.</summary>
<description>

All checked operands and bounds must be finite; NaN or either infinity reports Error
during active evaluation.

Numeric diagnostics use the formatter's default six significant digits; rounding affects
the message only, not the comparison.

</description>
*)
{endregion}
FUNCTION_BLOCK AssertNotEqual_LReal EXTENDS AssertionBase
VAR_INPUT
    IN : LREAL; //! Actual value checked or observed by this Assertion.
    Expected : LREAL; //! Value that must differ from IN under this Assertion's comparison rules.
END_VAR

SUPER^();

{region 'Documentation'}
(*!
<summary>Check inequality with the forbidden LREAL value.</summary>
*)
{endregion}
METHOD PROTECTED Assert
VAR
    Message : STRING(GVL_Constants.MessageLength);
    ExpectedText : STRING(GVL_Constants.AssertionValueLength);
    ActualText : STRING(GVL_Constants.AssertionValueLength);
END_VAR
IF NOT EvaluationActive THEN
    RETURN;
END_IF;

IF Result = E_Result.Error THEN
    RETURN;
END_IF;

IF NOT Tc2_Utilities.LrealIsFinite(x := IN) THEN
    Error(Message := 'Assertion error: IN must be finite.');
    RETURN;
END_IF;

IF NOT Tc2_Utilities.LrealIsFinite(x := Expected) THEN
    Error(Message := 'Assertion error: Expected must be finite.');
    RETURN;
END_IF;

IF Result = E_Result.Failed THEN
    RETURN;
END_IF;

IF IN = Expected THEN
    ExpectedText := CreateAssertionTextValue_LReal(Value := Expected);
    ActualText := CreateAssertionTextValue_LReal(Value := IN);
    Message := CONCAT('Assertion failed: values are equal but should differ. NotExpected = ',
        ExpectedText);
    Message := CONCAT(Message, ', Actual = ');
    Message := CONCAT(Message, ActualText);
    Message := CONCAT(Message, '.');
    Fail(Message := Message);
    RETURN;
END_IF;

Pass();
END_METHOD

END_FUNCTION_BLOCK

// ---- Framework/Assertions/POU/BasicTypes/LReal/AssertLessThan_LReal.TcPOU
{region 'Documentation'}
(*!
<summary>Check that IN is less than Maximum.</summary>
<description>

All checked operands and bounds must be finite; NaN or either infinity reports Error
during active evaluation.

Numeric diagnostics use the formatter's default six significant digits; rounding affects
the message only, not the comparison.

</description>
*)
{endregion}
FUNCTION_BLOCK AssertLessThan_LReal EXTENDS AssertionBase
VAR_INPUT
    IN : LREAL; //! Actual value checked or observed by this Assertion.
    Maximum : LREAL; //! Exclusive upper bound; the actual value or count must be smaller.
END_VAR

SUPER^();

{region 'Documentation'}
(*!
<summary>Check that IN is less than Maximum.</summary>
*)
{endregion}
METHOD PROTECTED Assert
VAR
    Message : STRING(GVL_Constants.MessageLength);
    MaximumText : STRING(GVL_Constants.AssertionValueLength);
    ActualText : STRING(GVL_Constants.AssertionValueLength);
END_VAR
IF NOT EvaluationActive THEN
    RETURN;
END_IF;

IF Result = E_Result.Error THEN
    RETURN;
END_IF;

IF NOT Tc2_Utilities.LrealIsFinite(x := IN) THEN
    Error(Message := 'Assertion error: IN must be finite.');
    RETURN;
END_IF;

IF NOT Tc2_Utilities.LrealIsFinite(x := Maximum) THEN
    Error(Message := 'Assertion error: Maximum must be finite.');
    RETURN;
END_IF;

IF Result = E_Result.Failed THEN
    RETURN;
END_IF;

IF IN >= Maximum THEN
    MaximumText := CreateAssertionTextValue_LReal(Value := Maximum);
    ActualText := CreateAssertionTextValue_LReal(Value := IN);
    Message := CONCAT('Assertion failed: value is not less than maximum. Maximum = ',
        MaximumText);
    Message := CONCAT(Message, ', Actual = ');
    Message := CONCAT(Message, ActualText);
    Message := CONCAT(Message, '.');
    Fail(Message := Message);
    RETURN;
END_IF;

Pass();
END_METHOD

END_FUNCTION_BLOCK

// ---- Framework/Assertions/POU/BasicTypes/LReal/AssertLessEqual_LReal.TcPOU
{region 'Documentation'}
(*!
<summary>Check that IN is at most Maximum.</summary>
<description>

All checked operands and bounds must be finite; NaN or either infinity reports Error
during active evaluation.

Numeric diagnostics use the formatter's default six significant digits; rounding affects
the message only, not the comparison.

</description>
*)
{endregion}
FUNCTION_BLOCK AssertLessEqual_LReal EXTENDS AssertionBase
VAR_INPUT
    IN : LREAL; //! Actual value checked or observed by this Assertion.
    Maximum : LREAL; //! Inclusive upper bound of the comparison; for a range, must not be below Minimum.
END_VAR

SUPER^();

{region 'Documentation'}
(*!
<summary>Check that IN is at most Maximum.</summary>
*)
{endregion}
METHOD PROTECTED Assert
VAR
    Message : STRING(GVL_Constants.MessageLength);
    MaximumText : STRING(GVL_Constants.AssertionValueLength);
    ActualText : STRING(GVL_Constants.AssertionValueLength);
END_VAR
IF NOT EvaluationActive THEN
    RETURN;
END_IF;

IF Result = E_Result.Error THEN
    RETURN;
END_IF;

IF NOT Tc2_Utilities.LrealIsFinite(x := IN) THEN
    Error(Message := 'Assertion error: IN must be finite.');
    RETURN;
END_IF;

IF NOT Tc2_Utilities.LrealIsFinite(x := Maximum) THEN
    Error(Message := 'Assertion error: Maximum must be finite.');
    RETURN;
END_IF;

IF Result = E_Result.Failed THEN
    RETURN;
END_IF;

IF IN > Maximum THEN
    MaximumText := CreateAssertionTextValue_LReal(Value := Maximum);
    ActualText := CreateAssertionTextValue_LReal(Value := IN);
    Message := CONCAT('Assertion failed: value is above maximum. Maximum = ',
        MaximumText);
    Message := CONCAT(Message, ', Actual = ');
    Message := CONCAT(Message, ActualText);
    Message := CONCAT(Message, '.');
    Fail(Message := Message);
    RETURN;
END_IF;

Pass();
END_METHOD

END_FUNCTION_BLOCK

// ---- Framework/Assertions/POU/BasicTypes/LReal/AssertGreaterThan_LReal.TcPOU
{region 'Documentation'}
(*!
<summary>Check that IN is greater than Minimum.</summary>
<description>

All checked operands and bounds must be finite; NaN or either infinity reports Error
during active evaluation.

Numeric diagnostics use the formatter's default six significant digits; rounding affects
the message only, not the comparison.

</description>
*)
{endregion}
FUNCTION_BLOCK AssertGreaterThan_LReal EXTENDS AssertionBase
VAR_INPUT
    IN : LREAL; //! Actual value checked or observed by this Assertion.
    Minimum : LREAL; //! Exclusive lower bound; the actual value or count must be greater.
END_VAR

SUPER^();

{region 'Documentation'}
(*!
<summary>Check that IN is greater than Minimum.</summary>
*)
{endregion}
METHOD PROTECTED Assert
VAR
    Message : STRING(GVL_Constants.MessageLength);
    MinimumText : STRING(GVL_Constants.AssertionValueLength);
    ActualText : STRING(GVL_Constants.AssertionValueLength);
END_VAR
IF NOT EvaluationActive THEN
    RETURN;
END_IF;

IF Result = E_Result.Error THEN
    RETURN;
END_IF;

IF NOT Tc2_Utilities.LrealIsFinite(x := IN) THEN
    Error(Message := 'Assertion error: IN must be finite.');
    RETURN;
END_IF;

IF NOT Tc2_Utilities.LrealIsFinite(x := Minimum) THEN
    Error(Message := 'Assertion error: Minimum must be finite.');
    RETURN;
END_IF;

IF Result = E_Result.Failed THEN
    RETURN;
END_IF;

IF IN <= Minimum THEN
    MinimumText := CreateAssertionTextValue_LReal(Value := Minimum);
    ActualText := CreateAssertionTextValue_LReal(Value := IN);
    Message := CONCAT('Assertion failed: value is not greater than minimum. Minimum = ',
        MinimumText);
    Message := CONCAT(Message, ', Actual = ');
    Message := CONCAT(Message, ActualText);
    Message := CONCAT(Message, '.');
    Fail(Message := Message);
    RETURN;
END_IF;

Pass();
END_METHOD

END_FUNCTION_BLOCK

// ---- Framework/Assertions/POU/BasicTypes/LReal/AssertGreaterEqual_LReal.TcPOU
{region 'Documentation'}
(*!
<summary>Check that IN is at least Minimum.</summary>
<description>

All checked operands and bounds must be finite; NaN or either infinity reports Error
during active evaluation.

Numeric diagnostics use the formatter's default six significant digits; rounding affects
the message only, not the comparison.

</description>
*)
{endregion}
FUNCTION_BLOCK AssertGreaterEqual_LReal EXTENDS AssertionBase
VAR_INPUT
    IN : LREAL; //! Actual value checked or observed by this Assertion.
    Minimum : LREAL; //! Inclusive lower bound of the comparison; for a range, must not exceed Maximum.
END_VAR

SUPER^();

{region 'Documentation'}
(*!
<summary>Check that IN is at least Minimum.</summary>
*)
{endregion}
METHOD PROTECTED Assert
VAR
    Message : STRING(GVL_Constants.MessageLength);
    MinimumText : STRING(GVL_Constants.AssertionValueLength);
    ActualText : STRING(GVL_Constants.AssertionValueLength);
END_VAR
IF NOT EvaluationActive THEN
    RETURN;
END_IF;

IF Result = E_Result.Error THEN
    RETURN;
END_IF;

IF NOT Tc2_Utilities.LrealIsFinite(x := IN) THEN
    Error(Message := 'Assertion error: IN must be finite.');
    RETURN;
END_IF;

IF NOT Tc2_Utilities.LrealIsFinite(x := Minimum) THEN
    Error(Message := 'Assertion error: Minimum must be finite.');
    RETURN;
END_IF;

IF Result = E_Result.Failed THEN
    RETURN;
END_IF;

IF IN < Minimum THEN
    MinimumText := CreateAssertionTextValue_LReal(Value := Minimum);
    ActualText := CreateAssertionTextValue_LReal(Value := IN);
    Message := CONCAT('Assertion failed: value is below minimum. Minimum = ',
        MinimumText);
    Message := CONCAT(Message, ', Actual = ');
    Message := CONCAT(Message, ActualText);
    Message := CONCAT(Message, '.');
    Fail(Message := Message);
    RETURN;
END_IF;

Pass();
END_METHOD

END_FUNCTION_BLOCK

// ---- Framework/Assertions/POU/BasicTypes/LReal/AssertInRange_LReal.TcPOU
{region 'Documentation'}
(*!
<summary>Checks whether the LREAL value is inside the inclusive range.</summary>
<description>

Minimum &gt; Maximum reports Error during active evaluation; equal bounds are
valid.

All checked operands and bounds must be finite; NaN or either infinity reports Error
during active evaluation.

Numeric diagnostics use the formatter's default six significant digits; rounding affects
the message only, not the comparison.

</description>
*)
{endregion}
FUNCTION_BLOCK AssertInRange_LReal EXTENDS AssertionBase
VAR_INPUT
    IN : LREAL; //! Actual value checked or observed by this Assertion.
    Minimum : LREAL; //! Inclusive lower bound of the comparison; for a range, must not exceed Maximum.
    Maximum : LREAL; //! Inclusive upper bound of the comparison; for a range, must not be below Minimum.
END_VAR

SUPER^();

{region 'Documentation'}
(*!
<summary>Check whether the LREAL value is inside the inclusive range.</summary>
*)
{endregion}
METHOD PROTECTED Assert
VAR
    Message : STRING(GVL_Constants.MessageLength);
    MinimumText : STRING(GVL_Constants.AssertionValueLength);
    MaximumText : STRING(GVL_Constants.AssertionValueLength);
    ActualText : STRING(GVL_Constants.AssertionValueLength);
END_VAR
IF NOT EvaluationActive THEN
    RETURN;
END_IF;

IF Result = E_Result.Error THEN
    RETURN;
END_IF;

IF NOT Tc2_Utilities.LrealIsFinite(x := IN) THEN
    Error(Message := 'Assertion error: IN must be finite.');
    RETURN;
END_IF;

IF NOT Tc2_Utilities.LrealIsFinite(x := Minimum) THEN
    Error(Message := 'Assertion error: Minimum must be finite.');
    RETURN;
END_IF;

IF NOT Tc2_Utilities.LrealIsFinite(x := Maximum) THEN
    Error(Message := 'Assertion error: Maximum must be finite.');
    RETURN;
END_IF;

IF Minimum > Maximum THEN
    MinimumText := CreateAssertionTextValue_LReal(Value := Minimum);
    MaximumText := CreateAssertionTextValue_LReal(Value := Maximum);
    Message := CONCAT('Assertion error: minimum exceeds maximum. Minimum = ',
        MinimumText);
    Message := CONCAT(Message, ', Maximum = ');
    Message := CONCAT(Message, MaximumText);
    Message := CONCAT(Message, '.');
    Error(Message := Message);
    RETURN;
END_IF;

IF Result = E_Result.Failed THEN
    RETURN;
END_IF;

IF (IN < Minimum) OR (IN > Maximum) THEN
    MinimumText := CreateAssertionTextValue_LReal(Value := Minimum);
    MaximumText := CreateAssertionTextValue_LReal(Value := Maximum);
    ActualText := CreateAssertionTextValue_LReal(Value := IN);
    Message := CONCAT('Assertion failed: value is outside allowed range. Minimum = ',
        MinimumText);
    Message := CONCAT(Message, ', Maximum = ');
    Message := CONCAT(Message, MaximumText);
    Message := CONCAT(Message, ', Actual = ');
    Message := CONCAT(Message, ActualText);
    Message := CONCAT(Message, '.');
    Fail(Message := Message);
    RETURN;
END_IF;

Pass();
END_METHOD

END_FUNCTION_BLOCK

// ---- Framework/Assertions/POU/BasicTypes/LReal/AssertNotInRange_LReal.TcPOU
{region 'Documentation'}
(*!
<summary>Checks whether the LREAL value is outside the inclusive range.</summary>
<description>

Minimum &gt; Maximum reports Error during active evaluation; equal bounds are
valid.

All checked operands and bounds must be finite; NaN or either infinity reports Error
during active evaluation.

Numeric diagnostics use the formatter's default six significant digits; rounding affects
the message only, not the comparison.

</description>
*)
{endregion}
FUNCTION_BLOCK AssertNotInRange_LReal EXTENDS AssertionBase
VAR_INPUT
    IN : LREAL; //! Actual value checked or observed by this Assertion.
    Minimum : LREAL; //! Inclusive lower bound of the comparison; for a range, must not exceed Maximum.
    Maximum : LREAL; //! Inclusive upper bound of the comparison; for a range, must not be below Minimum.
END_VAR

SUPER^();

{region 'Documentation'}
(*!
<summary>Check whether the LREAL value is outside the inclusive range.</summary>
*)
{endregion}
METHOD PROTECTED Assert
VAR
    Message : STRING(GVL_Constants.MessageLength);
    MinimumText : STRING(GVL_Constants.AssertionValueLength);
    MaximumText : STRING(GVL_Constants.AssertionValueLength);
    ActualText : STRING(GVL_Constants.AssertionValueLength);
END_VAR
IF NOT EvaluationActive THEN
    RETURN;
END_IF;

IF Result = E_Result.Error THEN
    RETURN;
END_IF;

IF NOT Tc2_Utilities.LrealIsFinite(x := IN) THEN
    Error(Message := 'Assertion error: IN must be finite.');
    RETURN;
END_IF;

IF NOT Tc2_Utilities.LrealIsFinite(x := Minimum) THEN
    Error(Message := 'Assertion error: Minimum must be finite.');
    RETURN;
END_IF;

IF NOT Tc2_Utilities.LrealIsFinite(x := Maximum) THEN
    Error(Message := 'Assertion error: Maximum must be finite.');
    RETURN;
END_IF;

IF Minimum > Maximum THEN
    MinimumText := CreateAssertionTextValue_LReal(Value := Minimum);
    MaximumText := CreateAssertionTextValue_LReal(Value := Maximum);
    Message := CONCAT('Assertion error: minimum exceeds maximum. Minimum = ',
        MinimumText);
    Message := CONCAT(Message, ', Maximum = ');
    Message := CONCAT(Message, MaximumText);
    Message := CONCAT(Message, '.');
    Error(Message := Message);
    RETURN;
END_IF;

IF Result = E_Result.Failed THEN
    RETURN;
END_IF;

IF (IN >= Minimum) AND (IN <= Maximum) THEN
    MinimumText := CreateAssertionTextValue_LReal(Value := Minimum);
    MaximumText := CreateAssertionTextValue_LReal(Value := Maximum);
    ActualText := CreateAssertionTextValue_LReal(Value := IN);
    Message := CONCAT('Assertion failed: value is inside forbidden range. Minimum = ',
        MinimumText);
    Message := CONCAT(Message, ', Maximum = ');
    Message := CONCAT(Message, MaximumText);
    Message := CONCAT(Message, ', Actual = ');
    Message := CONCAT(Message, ActualText);
    Message := CONCAT(Message, '.');
    Fail(Message := Message);
    RETURN;
END_IF;

Pass();
END_METHOD

END_FUNCTION_BLOCK

// ---- SelfTests/TestCases/TestSuite_AssertionFloatingPoint/Test_AssertionNonFinite_Real.TcPOU
{region 'Documentation'}
(*!
<summary>Checks REAL non-finite scalar operands and Error above held Failed.</summary>
<description>
Quiet NaN and both infinities are built by bit representation, never exceptional arithmetic.
Actual, expected/bound and tolerance roles are exercised separately across algorithm families.
NaNAfterFailure deliberately retains the preceding subject results; other rows reset them.
A disabled preparation call consumes subject resets before the next enabled observation.
Only outer checking Assertions contribute to the Test Case result.
Expected outcomes are explicit; production processing is inherited, not mirrored.
</description>
*)
{endregion}
FUNCTION_BLOCK Test_AssertionNonFinite_Real EXTENDS TestCaseBase
VAR
    FEqualSubject : AssertEqual_Real;
    FLessThanSubject : AssertLessThan_Real;
    FInRangeSubject : AssertInRange_Real;
    FEqualToleranceSubject : AssertEqualTolerance_Real;
    FNotEqualToleranceSubject : AssertNotEqualTolerance_Real;
    FActual : REAL;
    FExpected : REAL;
    FLower : REAL;
    FUpper : REAL;
    FTolerance : REAL;
    FQuietNaN : FloatingPointBits_Real;
    FPositiveInfinity : FloatingPointBits_Real;
    FNegativeInfinity : FloatingPointBits_Real;
    FExpectedEqualResult : E_Result;
    FExpectedLessThanResult : E_Result;
    FExpectedInRangeResult : E_Result;
    FExpectedEqualToleranceResult : E_Result;
    FExpectedNotEqualToleranceResult : E_Result;
    FExpectedFindings : UDINT;
    FCapture : EventBuffer;
    FEvents : ARRAY[1..CaptureLength] OF ST_Event;
    FCaptureFifo : ST_FifoStatus;
    FCaptureStatus : ST_EventBufferStatus;
    FRow : UINT;
    FRowPrepared : BOOL;
    FPreserveResults : BOOL;
    FObservationReady : BOOL;
    FChecked : BOOL;
    FSetupValid : BOOL;
END_VAR
VAR
    FEqualResult : AssertTrue;
    FEqualResultMatches : BOOL;
    FLessThanResult : AssertTrue;
    FLessThanResultMatches : BOOL;
    FInRangeResult : AssertTrue;
    FInRangeResultMatches : BOOL;
    FEqualToleranceResult : AssertTrue;
    FEqualToleranceResultMatches : BOOL;
    FNotEqualToleranceResult : AssertTrue;
    FNotEqualToleranceResultMatches : BOOL;
    FCaptureIntegrity : AssertTrue;
    FCaptureIntegrityMatches : BOOL;
    FFindingDetails : AssertTrue;
    FFindingDetailsMatch : BOOL;
END_VAR
VAR CONSTANT
    CaptureLength : UINT := 16;
    FixtureSize : UINT := 4;
    OneBits : DWORD := DWORD#16#3F800000;
    QuietNaNBits : DWORD := DWORD#16#7FC00000;
    PositiveInfinityBits : DWORD := DWORD#16#7F800000;
    NegativeInfinityBits : DWORD := DWORD#16#FF800000;
    ActualQuietNaN : UINT := 1;
    ActualPositiveInfinity : UINT := 2;
    ActualNegativeInfinity : UINT := 3;
    ExpectedQuietNaN : UINT := 4;
    ExpectedPositiveInfinity : UINT := 5;
    ExpectedNegativeInfinity : UINT := 6;
    LowerBoundQuietNaN : UINT := 7;
    LowerBoundPositiveInfinity : UINT := 8;
    LowerBoundNegativeInfinity : UINT := 9;
    UpperBoundQuietNaN : UINT := 10;
    UpperBoundPositiveInfinity : UINT := 11;
    UpperBoundNegativeInfinity : UINT := 12;
    ToleranceQuietNaN : UINT := 13;
    TolerancePositiveInfinity : UINT := 14;
    ToleranceNegativeInfinity : UINT := 15;
    FailureBeforeNaN : UINT := 16;
    NaNAfterFailure : UINT := 17;
    LastRow : UINT := NaNAfterFailure;
END_VAR

SUPER^();

{region 'Documentation'}
(*!
<summary>Collects only outer checking Assertions, never intentional subject findings.</summary>
*)
{endregion}
METHOD PROTECTED AggregateResults
VAR_INPUT
    Aggregator : I_ResultAggregator; //! Borrowed result sink owned by the outer Test Case; add this test's checking Assertions without resetting or retaining the sink.
END_VAR
Aggregator.AddProvider(Provider := FEqualResult);
Aggregator.AddProvider(Provider := FLessThanResult);
Aggregator.AddProvider(Provider := FInRangeResult);
Aggregator.AddProvider(Provider := FEqualToleranceResult);
Aggregator.AddProvider(Provider := FNotEqualToleranceResult);
Aggregator.AddProvider(Provider := FCaptureIntegrity);
Aggregator.AddProvider(Provider := FFindingDetails);
END_METHOD

{region 'Documentation'}
(*!
<summary>Calls each inherited production Assertion once using the selected row.</summary>
*)
{endregion}
METHOD PRIVATE CallSubjects
VAR_INPUT
    Enable : BOOL; //! Observation-enable input forwarded to the controlled Assertion subjects for this call.
END_VAR
FEqualSubject(Enable := Enable,
    State := E_State.Running,
    IN := FActual,
    Expected := FExpected);
FLessThanSubject(Enable := Enable,
    State := E_State.Running,
    IN := FActual,
    Maximum := FExpected);
FInRangeSubject(Enable := Enable,
    State := E_State.Running,
    IN := FActual,
    Minimum := FLower,
    Maximum := FUpper);
FEqualToleranceSubject(Enable := Enable,
    State := E_State.Running,
    IN := FActual,
    Expected := FExpected,
    Tolerance := FTolerance);
FNotEqualToleranceSubject(Enable := Enable,
    State := E_State.Running,
    IN := FActual,
    Expected := FExpected,
    Tolerance := FTolerance);
END_METHOD

{region 'Documentation'}
(*!
<summary>Extends base validation with subject and checking-Assertion setup.</summary>
*)
{endregion}
METHOD PROTECTED CheckInitialization : BOOL //! TRUE when the inherited initialization check and this concrete fixture check both accept the setup.
CheckInitialization := SUPER^.CheckInitialization();
IF NOT CheckInitialization THEN
    RETURN;
END_IF;

CheckInitialization := FSetupValid
    AND FEqualResult.IsInitialized
    AND FLessThanResult.IsInitialized
    AND FInRangeResult.IsInitialized
    AND FEqualToleranceResult.IsInitialized
    AND FNotEqualToleranceResult.IsInitialized
    AND FCaptureIntegrity.IsInitialized
    AND FFindingDetails.IsInitialized;
IF NOT CheckInitialization THEN
    EventPublisher.PublishEvent(Event := CreateFrameworkEvent(Name := Name,
        ResourceName := '',
        State := State,
        Severity := E_EventSeverity.Error,
        Message := 'Floating-point selftest setup or fixture representation failed.'));
END_IF;
END_METHOD

{region 'Documentation'}
(*!
<summary>Checks literal results and the ordered isolated findings from this row.</summary>
*)
{endregion}
METHOD PRIVATE CheckResults
VAR
    FindingIndex : UINT;
    FindingMatches : BOOL;
END_VAR
FEqualResultMatches := FEqualSubject.Result = FExpectedEqualResult;
FLessThanResultMatches := FLessThanSubject.Result = FExpectedLessThanResult;
FInRangeResultMatches := FInRangeSubject.Result = FExpectedInRangeResult;
FEqualToleranceResultMatches := FEqualToleranceSubject.Result = FExpectedEqualToleranceResult;
FNotEqualToleranceResultMatches := FNotEqualToleranceSubject.Result = FExpectedNotEqualToleranceResult;
FCaptureIntegrityMatches := (FCaptureStatus.SequenceId = FExpectedFindings)
    AND (FCaptureStatus.LostEventCount = 0);

FindingIndex := 1;
FFindingDetailsMatch := TRUE;
IF (FExpectedEqualResult = E_Result.Failed) OR (FExpectedEqualResult = E_Result.Error) THEN
    FindingMatches := IsFindingValid(Index := FindingIndex,
        ExpectedName := FEqualSubject.Name,
        ExpectedResult := FExpectedEqualResult);
    FFindingDetailsMatch := FFindingDetailsMatch AND FindingMatches;
    FindingIndex := FindingIndex + 1;
END_IF;
IF (FExpectedLessThanResult = E_Result.Failed) OR (FExpectedLessThanResult = E_Result.Error) THEN
    FindingMatches := IsFindingValid(Index := FindingIndex,
        ExpectedName := FLessThanSubject.Name,
        ExpectedResult := FExpectedLessThanResult);
    FFindingDetailsMatch := FFindingDetailsMatch AND FindingMatches;
    FindingIndex := FindingIndex + 1;
END_IF;
IF (FExpectedInRangeResult = E_Result.Failed) OR (FExpectedInRangeResult = E_Result.Error) THEN
    FindingMatches := IsFindingValid(Index := FindingIndex,
        ExpectedName := FInRangeSubject.Name,
        ExpectedResult := FExpectedInRangeResult);
    FFindingDetailsMatch := FFindingDetailsMatch AND FindingMatches;
    FindingIndex := FindingIndex + 1;
END_IF;
IF (FExpectedEqualToleranceResult = E_Result.Failed) OR (FExpectedEqualToleranceResult = E_Result.Error) THEN
    FindingMatches := IsFindingValid(Index := FindingIndex,
        ExpectedName := FEqualToleranceSubject.Name,
        ExpectedResult := FExpectedEqualToleranceResult);
    FFindingDetailsMatch := FFindingDetailsMatch AND FindingMatches;
    FindingIndex := FindingIndex + 1;
END_IF;
IF (FExpectedNotEqualToleranceResult = E_Result.Failed) OR (FExpectedNotEqualToleranceResult = E_Result.Error) THEN
    FindingMatches := IsFindingValid(Index := FindingIndex,
        ExpectedName := FNotEqualToleranceSubject.Name,
        ExpectedResult := FExpectedNotEqualToleranceResult);
    FFindingDetailsMatch := FFindingDetailsMatch AND FindingMatches;
    FindingIndex := FindingIndex + 1;
END_IF;
END_METHOD

{region 'Documentation'}
(*!
<summary>Configures checking Assertions; subject actions remain in the test script.</summary>
*)
{endregion}
METHOD PROTECTED Configure
VAR
    Initialized : BOOL;
END_VAR
FPreparationStateCount := 0;
FTestStateCount := 1;
FSetupValid := InitializeValues();
FEqualResult.Initialize(Parent := THIS^,
    AssertionName := 'EqualResult');
FLessThanResult.Initialize(Parent := THIS^,
    AssertionName := 'LessThanResult');
FInRangeResult.Initialize(Parent := THIS^,
    AssertionName := 'InRangeResult');
FEqualToleranceResult.Initialize(Parent := THIS^,
    AssertionName := 'EqualToleranceResult');
FNotEqualToleranceResult.Initialize(Parent := THIS^,
    AssertionName := 'NotEqualToleranceResult');
FCaptureIntegrity.Initialize(Parent := THIS^,
    AssertionName := 'CaptureIntegrity');
FFindingDetails.Initialize(Parent := THIS^,
    AssertionName := 'FindingDetails');
Initialized := FCapture.Initialize(Buffer := FEvents,
    FifoControl := FCaptureFifo,
    Status := FCaptureStatus);
FSetupValid := FSetupValid AND Initialized;
FEqualSubject.BindPublisher(Publisher := FCapture);
Initialized := FEqualSubject.Initialize(Parent := THIS^,
    AssertionName := 'EqualSubject');
FSetupValid := FSetupValid AND Initialized;
FLessThanSubject.BindPublisher(Publisher := FCapture);
Initialized := FLessThanSubject.Initialize(Parent := THIS^,
    AssertionName := 'LessThanSubject');
FSetupValid := FSetupValid AND Initialized;
FInRangeSubject.BindPublisher(Publisher := FCapture);
Initialized := FInRangeSubject.Initialize(Parent := THIS^,
    AssertionName := 'InRangeSubject');
FSetupValid := FSetupValid AND Initialized;
FEqualToleranceSubject.BindPublisher(Publisher := FCapture);
Initialized := FEqualToleranceSubject.Initialize(Parent := THIS^,
    AssertionName := 'EqualToleranceSubject');
FSetupValid := FSetupValid AND Initialized;
FNotEqualToleranceSubject.BindPublisher(Publisher := FCapture);
Initialized := FNotEqualToleranceSubject.Initialize(Parent := THIS^,
    AssertionName := 'NotEqualToleranceSubject');
FSetupValid := FSetupValid AND Initialized;
END_METHOD

{region 'Documentation'}
(*!
<summary>Establishes typed fixtures and verifies their representation before any subject call.</summary>
*)
{endregion}
METHOD PRIVATE InitializeValues : BOOL //! TRUE when fixture sizes and floating-point bit representations match their explicit expected patterns.
VAR
    Representation : FloatingPointBits_Real;
END_VAR
Representation.Value := REAL#1.0;
InitializeValues := (SIZEOF(Representation) = FixtureSize)
    AND (Representation.Bits = OneBits);

FQuietNaN.Bits := QuietNaNBits;
Representation.Value := FQuietNaN.Value;
InitializeValues := InitializeValues AND (Representation.Bits = QuietNaNBits);
FPositiveInfinity.Bits := PositiveInfinityBits;
Representation.Value := FPositiveInfinity.Value;
InitializeValues := InitializeValues AND (Representation.Bits = PositiveInfinityBits);
FNegativeInfinity.Bits := NegativeInfinityBits;
Representation.Value := FNegativeInfinity.Value;
InitializeValues := InitializeValues AND (Representation.Bits = NegativeInfinityBits);
END_METHOD

{region 'Documentation'}
(*!
<summary>Reads a captured finding; the caller bounds the index by 5 subjects.</summary>
*)
{endregion}
METHOD PRIVATE IsFindingValid : BOOL //! TRUE when the selected captured finding satisfies the scenario metadata and diagnostic checks.
VAR_INPUT
    Index : UINT; //! One-based index in the retained isolated event capture.
    ExpectedName : STRING(GVL_Constants.NameLength); //! Independently authored Assertion name expected in the selected finding.
    ExpectedResult : E_Result; //! Independently authored finding result.
END_VAR
IsFindingValid := (FEvents[Index].SequenceId = UINT_TO_UDINT(Index))
    AND (FEvents[Index].Name = ExpectedName)
    AND (FEvents[Index].OwnerScope = E_OwnerScope.Assertion)
    AND (FEvents[Index].EventType = E_EventType.Result)
    AND (FEvents[Index].State = E_State.Running)
    AND (FEvents[Index].Result = ExpectedResult)
    AND (FEvents[Index].Message <> '');
END_METHOD

{region 'Documentation'}
(*!
<summary>Completes abort without asynchronous resources.</summary>
*)
{endregion}
METHOD PROTECTED ProcessAbort
VAR_INPUT
    Enable : BOOL; //! Phase permission supplied by the owning Test Case; FALSE does not authorize progression, while observation may continue.
END_VAR
IF Enable THEN
    CompleteAbort();
END_IF;
END_METHOD

{region 'Documentation'}
(*!
<summary>Latches checked observations before the next script step may proceed.</summary>
*)
{endregion}
METHOD PROTECTED ProcessAssertions
VAR_INPUT
    Enable : BOOL; //! Phase permission supplied by the owning Test Case; FALSE does not authorize progression, while observation may continue.
END_VAR
VAR
    Evaluate : BOOL;
END_VAR
Evaluate := Enable AND FObservationReady;
FEqualResult(Enable := Evaluate,
    State := State,
    IN := FEqualResultMatches);
FLessThanResult(Enable := Evaluate,
    State := State,
    IN := FLessThanResultMatches);
FInRangeResult(Enable := Evaluate,
    State := State,
    IN := FInRangeResultMatches);
FEqualToleranceResult(Enable := Evaluate,
    State := State,
    IN := FEqualToleranceResultMatches);
FNotEqualToleranceResult(Enable := Evaluate,
    State := State,
    IN := FNotEqualToleranceResultMatches);
FCaptureIntegrity(Enable := Evaluate,
    State := State,
    IN := FCaptureIntegrityMatches);
FFindingDetails(Enable := Evaluate,
    State := State,
    IN := FFindingDetailsMatch);
IF Evaluate THEN
    FChecked := TRUE;
END_IF;
END_METHOD

{region 'Documentation'}
(*!
<summary>No Preparation phase is required.</summary>
*)
{endregion}
METHOD PROTECTED ProcessPreparations
VAR_INPUT
    // SA0033: Required hook; this test has no Preparation phase.
    {attribute 'analysis' := '-33'}
    Enable : BOOL; //! Phase permission supplied by the owning Test Case; FALSE does not authorize progression, while observation may continue.
END_VAR
END_METHOD

{region 'Documentation'}
(*!
<summary>Restarts the script and resets the checking Assertions.</summary>
*)
{endregion}
METHOD PROTECTED ProcessReset
FRow := ActualQuietNaN;
FRowPrepared := FALSE;
FChecked := FALSE;
FObservationReady := FALSE;
FEqualResult.Reset();
FEqualResultMatches := TRUE;
FLessThanResult.Reset();
FLessThanResultMatches := TRUE;
FInRangeResult.Reset();
FInRangeResultMatches := TRUE;
FEqualToleranceResult.Reset();
FEqualToleranceResultMatches := TRUE;
FNotEqualToleranceResult.Reset();
FNotEqualToleranceResultMatches := TRUE;
FCaptureIntegrity.Reset();
FCaptureIntegrityMatches := TRUE;
FFindingDetails.Reset();
FFindingDetailsMatch := TRUE;
CompleteReset();
END_METHOD

{region 'Documentation'}
(*!
<summary>Advances one bounded script step per active PLC cycle.</summary>
*)
{endregion}
METHOD PROTECTED ProcessTests
VAR_INPUT
    Enable : BOOL; //! Phase permission supplied by the owning Test Case; FALSE does not authorize progression, while observation may continue.
END_VAR
IF NOT Enable THEN
    RETURN;
END_IF;

IF FChecked THEN
    FChecked := FALSE;
    FObservationReady := FALSE;
    IF FRow = LastRow THEN
        CompleteTests();
        RETURN;
    END_IF;
    FRow := FRow + 1;
    FRowPrepared := FALSE;
END_IF;

IF NOT FRowPrepared THEN
    SelectRow();
    FCapture.Reset();
    IF NOT FPreserveResults THEN
        ResetSubjects();
    END_IF;
    CallSubjects(Enable := FALSE);
    FRowPrepared := TRUE;
ELSE
    CallSubjects(Enable := TRUE);
    CheckResults();
    FObservationReady := TRUE;
END_IF;
END_METHOD

{region 'Documentation'}
(*!
<summary>Requests fresh subject results before the next disabled call.</summary>
*)
{endregion}
METHOD PRIVATE ResetSubjects
FEqualSubject.Reset();
FLessThanSubject.Reset();
FInRangeSubject.Reset();
FEqualToleranceSubject.Reset();
FNotEqualToleranceSubject.Reset();
END_METHOD

{region 'Documentation'}
(*!
<summary>Selects independent literal outcomes; only named escalation rows preserve results.</summary>
*)
{endregion}
METHOD PRIVATE SelectRow
FPreserveResults := FALSE;
CASE FRow OF
    ActualQuietNaN:
        FActual := FQuietNaN.Value;
        FExpected := REAL#1.0;
        FLower := REAL#0.0;
        FUpper := REAL#2.0;
        FTolerance := REAL#0.5;
        FExpectedEqualResult := E_Result.Error;
        FExpectedLessThanResult := E_Result.Error;
        FExpectedInRangeResult := E_Result.Error;
        FExpectedEqualToleranceResult := E_Result.Error;
        FExpectedNotEqualToleranceResult := E_Result.Error;
        FExpectedFindings := 5;
    ActualPositiveInfinity:
        FActual := FPositiveInfinity.Value;
        FExpected := REAL#1.0;
        FLower := REAL#0.0;
        FUpper := REAL#2.0;
        FTolerance := REAL#0.5;
        FExpectedEqualResult := E_Result.Error;
        FExpectedLessThanResult := E_Result.Error;
        FExpectedInRangeResult := E_Result.Error;
        FExpectedEqualToleranceResult := E_Result.Error;
        FExpectedNotEqualToleranceResult := E_Result.Error;
        FExpectedFindings := 5;
    ActualNegativeInfinity:
        FActual := FNegativeInfinity.Value;
        FExpected := REAL#1.0;
        FLower := REAL#0.0;
        FUpper := REAL#2.0;
        FTolerance := REAL#0.5;
        FExpectedEqualResult := E_Result.Error;
        FExpectedLessThanResult := E_Result.Error;
        FExpectedInRangeResult := E_Result.Error;
        FExpectedEqualToleranceResult := E_Result.Error;
        FExpectedNotEqualToleranceResult := E_Result.Error;
        FExpectedFindings := 5;
    ExpectedQuietNaN:
        FActual := REAL#1.0;
        FExpected := FQuietNaN.Value;
        FLower := REAL#0.0;
        FUpper := REAL#2.0;
        FTolerance := REAL#0.5;
        FExpectedEqualResult := E_Result.Error;
        FExpectedLessThanResult := E_Result.Error;
        FExpectedInRangeResult := E_Result.Passed;
        FExpectedEqualToleranceResult := E_Result.Error;
        FExpectedNotEqualToleranceResult := E_Result.Error;
        FExpectedFindings := 4;
    ExpectedPositiveInfinity:
        FActual := REAL#1.0;
        FExpected := FPositiveInfinity.Value;
        FLower := REAL#0.0;
        FUpper := REAL#2.0;
        FTolerance := REAL#0.5;
        FExpectedEqualResult := E_Result.Error;
        FExpectedLessThanResult := E_Result.Error;
        FExpectedInRangeResult := E_Result.Passed;
        FExpectedEqualToleranceResult := E_Result.Error;
        FExpectedNotEqualToleranceResult := E_Result.Error;
        FExpectedFindings := 4;
    ExpectedNegativeInfinity:
        FActual := REAL#1.0;
        FExpected := FNegativeInfinity.Value;
        FLower := REAL#0.0;
        FUpper := REAL#2.0;
        FTolerance := REAL#0.5;
        FExpectedEqualResult := E_Result.Error;
        FExpectedLessThanResult := E_Result.Error;
        FExpectedInRangeResult := E_Result.Passed;
        FExpectedEqualToleranceResult := E_Result.Error;
        FExpectedNotEqualToleranceResult := E_Result.Error;
        FExpectedFindings := 4;
    LowerBoundQuietNaN:
        FActual := REAL#1.0;
        FExpected := REAL#1.0;
        FLower := FQuietNaN.Value;
        FUpper := REAL#2.0;
        FTolerance := REAL#0.5;
        FExpectedEqualResult := E_Result.Passed;
        FExpectedLessThanResult := E_Result.Failed;
        FExpectedInRangeResult := E_Result.Error;
        FExpectedEqualToleranceResult := E_Result.Passed;
        FExpectedNotEqualToleranceResult := E_Result.Failed;
        FExpectedFindings := 3;
    LowerBoundPositiveInfinity:
        FActual := REAL#1.0;
        FExpected := REAL#1.0;
        FLower := FPositiveInfinity.Value;
        FUpper := REAL#2.0;
        FTolerance := REAL#0.5;
        FExpectedEqualResult := E_Result.Passed;
        FExpectedLessThanResult := E_Result.Failed;
        FExpectedInRangeResult := E_Result.Error;
        FExpectedEqualToleranceResult := E_Result.Passed;
        FExpectedNotEqualToleranceResult := E_Result.Failed;
        FExpectedFindings := 3;
    LowerBoundNegativeInfinity:
        FActual := REAL#1.0;
        FExpected := REAL#1.0;
        FLower := FNegativeInfinity.Value;
        FUpper := REAL#2.0;
        FTolerance := REAL#0.5;
        FExpectedEqualResult := E_Result.Passed;
        FExpectedLessThanResult := E_Result.Failed;
        FExpectedInRangeResult := E_Result.Error;
        FExpectedEqualToleranceResult := E_Result.Passed;
        FExpectedNotEqualToleranceResult := E_Result.Failed;
        FExpectedFindings := 3;
    UpperBoundQuietNaN:
        FActual := REAL#1.0;
        FExpected := REAL#1.0;
        FLower := REAL#0.0;
        FUpper := FQuietNaN.Value;
        FTolerance := REAL#0.5;
        FExpectedEqualResult := E_Result.Passed;
        FExpectedLessThanResult := E_Result.Failed;
        FExpectedInRangeResult := E_Result.Error;
        FExpectedEqualToleranceResult := E_Result.Passed;
        FExpectedNotEqualToleranceResult := E_Result.Failed;
        FExpectedFindings := 3;
    UpperBoundPositiveInfinity:
        FActual := REAL#1.0;
        FExpected := REAL#1.0;
        FLower := REAL#0.0;
        FUpper := FPositiveInfinity.Value;
        FTolerance := REAL#0.5;
        FExpectedEqualResult := E_Result.Passed;
        FExpectedLessThanResult := E_Result.Failed;
        FExpectedInRangeResult := E_Result.Error;
        FExpectedEqualToleranceResult := E_Result.Passed;
        FExpectedNotEqualToleranceResult := E_Result.Failed;
        FExpectedFindings := 3;
    UpperBoundNegativeInfinity:
        FActual := REAL#1.0;
        FExpected := REAL#1.0;
        FLower := REAL#0.0;
        FUpper := FNegativeInfinity.Value;
        FTolerance := REAL#0.5;
        FExpectedEqualResult := E_Result.Passed;
        FExpectedLessThanResult := E_Result.Failed;
        FExpectedInRangeResult := E_Result.Error;
        FExpectedEqualToleranceResult := E_Result.Passed;
        FExpectedNotEqualToleranceResult := E_Result.Failed;
        FExpectedFindings := 3;
    ToleranceQuietNaN:
        FActual := REAL#1.0;
        FExpected := REAL#1.0;
        FLower := REAL#0.0;
        FUpper := REAL#2.0;
        FTolerance := FQuietNaN.Value;
        FExpectedEqualResult := E_Result.Passed;
        FExpectedLessThanResult := E_Result.Failed;
        FExpectedInRangeResult := E_Result.Passed;
        FExpectedEqualToleranceResult := E_Result.Error;
        FExpectedNotEqualToleranceResult := E_Result.Error;
        FExpectedFindings := 3;
    TolerancePositiveInfinity:
        FActual := REAL#1.0;
        FExpected := REAL#1.0;
        FLower := REAL#0.0;
        FUpper := REAL#2.0;
        FTolerance := FPositiveInfinity.Value;
        FExpectedEqualResult := E_Result.Passed;
        FExpectedLessThanResult := E_Result.Failed;
        FExpectedInRangeResult := E_Result.Passed;
        FExpectedEqualToleranceResult := E_Result.Error;
        FExpectedNotEqualToleranceResult := E_Result.Error;
        FExpectedFindings := 3;
    ToleranceNegativeInfinity:
        FActual := REAL#1.0;
        FExpected := REAL#1.0;
        FLower := REAL#0.0;
        FUpper := REAL#2.0;
        FTolerance := FNegativeInfinity.Value;
        FExpectedEqualResult := E_Result.Passed;
        FExpectedLessThanResult := E_Result.Failed;
        FExpectedInRangeResult := E_Result.Passed;
        FExpectedEqualToleranceResult := E_Result.Error;
        FExpectedNotEqualToleranceResult := E_Result.Error;
        FExpectedFindings := 3;
    FailureBeforeNaN:
        FActual := REAL#3.0;
        FExpected := REAL#1.0;
        FLower := REAL#0.0;
        FUpper := REAL#2.0;
        FTolerance := REAL#0.5;
        FExpectedEqualResult := E_Result.Failed;
        FExpectedLessThanResult := E_Result.Failed;
        FExpectedInRangeResult := E_Result.Failed;
        FExpectedEqualToleranceResult := E_Result.Failed;
        FExpectedNotEqualToleranceResult := E_Result.Passed;
        FExpectedFindings := 4;
    NaNAfterFailure:
        FActual := FQuietNaN.Value;
        FExpected := REAL#1.0;
        FLower := REAL#0.0;
        FUpper := REAL#2.0;
        FTolerance := REAL#0.5;
        FExpectedEqualResult := E_Result.Error;
        FExpectedLessThanResult := E_Result.Error;
        FExpectedInRangeResult := E_Result.Error;
        FExpectedEqualToleranceResult := E_Result.Error;
        FExpectedNotEqualToleranceResult := E_Result.Error;
        FExpectedFindings := 5;
        FPreserveResults := TRUE;
ELSE
    Error(Message := 'Unknown floating-point test row.');
END_CASE;
END_METHOD

END_FUNCTION_BLOCK

// ---- SelfTests/TestCases/TestSuite_AssertionFloatingPoint/Test_AssertionNonFinite_LReal.TcPOU
{region 'Documentation'}
(*!
<summary>Checks LREAL non-finite scalar operands and Error above held Failed.</summary>
<description>
Quiet NaN and both infinities are built by bit representation, never exceptional arithmetic.
Actual, expected/bound and tolerance roles are exercised separately across algorithm families.
NaNAfterFailure deliberately retains the preceding subject results; other rows reset them.
A disabled preparation call consumes subject resets before the next enabled observation.
Only outer checking Assertions contribute to the Test Case result.
Expected outcomes are explicit; production processing is inherited, not mirrored.
</description>
*)
{endregion}
FUNCTION_BLOCK Test_AssertionNonFinite_LReal EXTENDS TestCaseBase
VAR
    FEqualSubject : AssertEqual_LReal;
    FLessThanSubject : AssertLessThan_LReal;
    FInRangeSubject : AssertInRange_LReal;
    FEqualToleranceSubject : AssertEqualTolerance_LReal;
    FNotEqualToleranceSubject : AssertNotEqualTolerance_LReal;
    FActual : LREAL;
    FExpected : LREAL;
    FLower : LREAL;
    FUpper : LREAL;
    FTolerance : LREAL;
    FQuietNaN : FloatingPointBits_LReal;
    FPositiveInfinity : FloatingPointBits_LReal;
    FNegativeInfinity : FloatingPointBits_LReal;
    FExpectedEqualResult : E_Result;
    FExpectedLessThanResult : E_Result;
    FExpectedInRangeResult : E_Result;
    FExpectedEqualToleranceResult : E_Result;
    FExpectedNotEqualToleranceResult : E_Result;
    FExpectedFindings : UDINT;
    FCapture : EventBuffer;
    FEvents : ARRAY[1..CaptureLength] OF ST_Event;
    FCaptureFifo : ST_FifoStatus;
    FCaptureStatus : ST_EventBufferStatus;
    FRow : UINT;
    FRowPrepared : BOOL;
    FPreserveResults : BOOL;
    FObservationReady : BOOL;
    FChecked : BOOL;
    FSetupValid : BOOL;
END_VAR
VAR
    FEqualResult : AssertTrue;
    FEqualResultMatches : BOOL;
    FLessThanResult : AssertTrue;
    FLessThanResultMatches : BOOL;
    FInRangeResult : AssertTrue;
    FInRangeResultMatches : BOOL;
    FEqualToleranceResult : AssertTrue;
    FEqualToleranceResultMatches : BOOL;
    FNotEqualToleranceResult : AssertTrue;
    FNotEqualToleranceResultMatches : BOOL;
    FCaptureIntegrity : AssertTrue;
    FCaptureIntegrityMatches : BOOL;
    FFindingDetails : AssertTrue;
    FFindingDetailsMatch : BOOL;
END_VAR
VAR CONSTANT
    CaptureLength : UINT := 16;
    FixtureSize : UINT := 8;
    OneBits : LWORD := LWORD#16#3FF0000000000000;
    QuietNaNBits : LWORD := LWORD#16#7FF8000000000000;
    PositiveInfinityBits : LWORD := LWORD#16#7FF0000000000000;
    NegativeInfinityBits : LWORD := LWORD#16#FFF0000000000000;
    ActualQuietNaN : UINT := 1;
    ActualPositiveInfinity : UINT := 2;
    ActualNegativeInfinity : UINT := 3;
    ExpectedQuietNaN : UINT := 4;
    ExpectedPositiveInfinity : UINT := 5;
    ExpectedNegativeInfinity : UINT := 6;
    LowerBoundQuietNaN : UINT := 7;
    LowerBoundPositiveInfinity : UINT := 8;
    LowerBoundNegativeInfinity : UINT := 9;
    UpperBoundQuietNaN : UINT := 10;
    UpperBoundPositiveInfinity : UINT := 11;
    UpperBoundNegativeInfinity : UINT := 12;
    ToleranceQuietNaN : UINT := 13;
    TolerancePositiveInfinity : UINT := 14;
    ToleranceNegativeInfinity : UINT := 15;
    FailureBeforeNaN : UINT := 16;
    NaNAfterFailure : UINT := 17;
    LastRow : UINT := NaNAfterFailure;
END_VAR

SUPER^();

{region 'Documentation'}
(*!
<summary>Collects only outer checking Assertions, never intentional subject findings.</summary>
*)
{endregion}
METHOD PROTECTED AggregateResults
VAR_INPUT
    Aggregator : I_ResultAggregator; //! Borrowed result sink owned by the outer Test Case; add this test's checking Assertions without resetting or retaining the sink.
END_VAR
Aggregator.AddProvider(Provider := FEqualResult);
Aggregator.AddProvider(Provider := FLessThanResult);
Aggregator.AddProvider(Provider := FInRangeResult);
Aggregator.AddProvider(Provider := FEqualToleranceResult);
Aggregator.AddProvider(Provider := FNotEqualToleranceResult);
Aggregator.AddProvider(Provider := FCaptureIntegrity);
Aggregator.AddProvider(Provider := FFindingDetails);
END_METHOD

{region 'Documentation'}
(*!
<summary>Calls each inherited production Assertion once using the selected row.</summary>
*)
{endregion}
METHOD PRIVATE CallSubjects
VAR_INPUT
    Enable : BOOL; //! Observation-enable input forwarded to the controlled Assertion subjects for this call.
END_VAR
FEqualSubject(Enable := Enable,
    State := E_State.Running,
    IN := FActual,
    Expected := FExpected);
FLessThanSubject(Enable := Enable,
    State := E_State.Running,
    IN := FActual,
    Maximum := FExpected);
FInRangeSubject(Enable := Enable,
    State := E_State.Running,
    IN := FActual,
    Minimum := FLower,
    Maximum := FUpper);
FEqualToleranceSubject(Enable := Enable,
    State := E_State.Running,
    IN := FActual,
    Expected := FExpected,
    Tolerance := FTolerance);
FNotEqualToleranceSubject(Enable := Enable,
    State := E_State.Running,
    IN := FActual,
    Expected := FExpected,
    Tolerance := FTolerance);
END_METHOD

{region 'Documentation'}
(*!
<summary>Extends base validation with subject and checking-Assertion setup.</summary>
*)
{endregion}
METHOD PROTECTED CheckInitialization : BOOL //! TRUE when the inherited initialization check and this concrete fixture check both accept the setup.
CheckInitialization := SUPER^.CheckInitialization();
IF NOT CheckInitialization THEN
    RETURN;
END_IF;

CheckInitialization := FSetupValid
    AND FEqualResult.IsInitialized
    AND FLessThanResult.IsInitialized
    AND FInRangeResult.IsInitialized
    AND FEqualToleranceResult.IsInitialized
    AND FNotEqualToleranceResult.IsInitialized
    AND FCaptureIntegrity.IsInitialized
    AND FFindingDetails.IsInitialized;
IF NOT CheckInitialization THEN
    EventPublisher.PublishEvent(Event := CreateFrameworkEvent(Name := Name,
        ResourceName := '',
        State := State,
        Severity := E_EventSeverity.Error,
        Message := 'Floating-point selftest setup or fixture representation failed.'));
END_IF;
END_METHOD

{region 'Documentation'}
(*!
<summary>Checks literal results and the ordered isolated findings from this row.</summary>
*)
{endregion}
METHOD PRIVATE CheckResults
VAR
    FindingIndex : UINT;
    FindingMatches : BOOL;
END_VAR
FEqualResultMatches := FEqualSubject.Result = FExpectedEqualResult;
FLessThanResultMatches := FLessThanSubject.Result = FExpectedLessThanResult;
FInRangeResultMatches := FInRangeSubject.Result = FExpectedInRangeResult;
FEqualToleranceResultMatches := FEqualToleranceSubject.Result = FExpectedEqualToleranceResult;
FNotEqualToleranceResultMatches := FNotEqualToleranceSubject.Result = FExpectedNotEqualToleranceResult;
FCaptureIntegrityMatches := (FCaptureStatus.SequenceId = FExpectedFindings)
    AND (FCaptureStatus.LostEventCount = 0);

FindingIndex := 1;
FFindingDetailsMatch := TRUE;
IF (FExpectedEqualResult = E_Result.Failed) OR (FExpectedEqualResult = E_Result.Error) THEN
    FindingMatches := IsFindingValid(Index := FindingIndex,
        ExpectedName := FEqualSubject.Name,
        ExpectedResult := FExpectedEqualResult);
    FFindingDetailsMatch := FFindingDetailsMatch AND FindingMatches;
    FindingIndex := FindingIndex + 1;
END_IF;
IF (FExpectedLessThanResult = E_Result.Failed) OR (FExpectedLessThanResult = E_Result.Error) THEN
    FindingMatches := IsFindingValid(Index := FindingIndex,
        ExpectedName := FLessThanSubject.Name,
        ExpectedResult := FExpectedLessThanResult);
    FFindingDetailsMatch := FFindingDetailsMatch AND FindingMatches;
    FindingIndex := FindingIndex + 1;
END_IF;
IF (FExpectedInRangeResult = E_Result.Failed) OR (FExpectedInRangeResult = E_Result.Error) THEN
    FindingMatches := IsFindingValid(Index := FindingIndex,
        ExpectedName := FInRangeSubject.Name,
        ExpectedResult := FExpectedInRangeResult);
    FFindingDetailsMatch := FFindingDetailsMatch AND FindingMatches;
    FindingIndex := FindingIndex + 1;
END_IF;
IF (FExpectedEqualToleranceResult = E_Result.Failed) OR (FExpectedEqualToleranceResult = E_Result.Error) THEN
    FindingMatches := IsFindingValid(Index := FindingIndex,
        ExpectedName := FEqualToleranceSubject.Name,
        ExpectedResult := FExpectedEqualToleranceResult);
    FFindingDetailsMatch := FFindingDetailsMatch AND FindingMatches;
    FindingIndex := FindingIndex + 1;
END_IF;
IF (FExpectedNotEqualToleranceResult = E_Result.Failed) OR (FExpectedNotEqualToleranceResult = E_Result.Error) THEN
    FindingMatches := IsFindingValid(Index := FindingIndex,
        ExpectedName := FNotEqualToleranceSubject.Name,
        ExpectedResult := FExpectedNotEqualToleranceResult);
    FFindingDetailsMatch := FFindingDetailsMatch AND FindingMatches;
    FindingIndex := FindingIndex + 1;
END_IF;
END_METHOD

{region 'Documentation'}
(*!
<summary>Configures checking Assertions; subject actions remain in the test script.</summary>
*)
{endregion}
METHOD PROTECTED Configure
VAR
    Initialized : BOOL;
END_VAR
FPreparationStateCount := 0;
FTestStateCount := 1;
FSetupValid := InitializeValues();
FEqualResult.Initialize(Parent := THIS^,
    AssertionName := 'EqualResult');
FLessThanResult.Initialize(Parent := THIS^,
    AssertionName := 'LessThanResult');
FInRangeResult.Initialize(Parent := THIS^,
    AssertionName := 'InRangeResult');
FEqualToleranceResult.Initialize(Parent := THIS^,
    AssertionName := 'EqualToleranceResult');
FNotEqualToleranceResult.Initialize(Parent := THIS^,
    AssertionName := 'NotEqualToleranceResult');
FCaptureIntegrity.Initialize(Parent := THIS^,
    AssertionName := 'CaptureIntegrity');
FFindingDetails.Initialize(Parent := THIS^,
    AssertionName := 'FindingDetails');
Initialized := FCapture.Initialize(Buffer := FEvents,
    FifoControl := FCaptureFifo,
    Status := FCaptureStatus);
FSetupValid := FSetupValid AND Initialized;
FEqualSubject.BindPublisher(Publisher := FCapture);
Initialized := FEqualSubject.Initialize(Parent := THIS^,
    AssertionName := 'EqualSubject');
FSetupValid := FSetupValid AND Initialized;
FLessThanSubject.BindPublisher(Publisher := FCapture);
Initialized := FLessThanSubject.Initialize(Parent := THIS^,
    AssertionName := 'LessThanSubject');
FSetupValid := FSetupValid AND Initialized;
FInRangeSubject.BindPublisher(Publisher := FCapture);
Initialized := FInRangeSubject.Initialize(Parent := THIS^,
    AssertionName := 'InRangeSubject');
FSetupValid := FSetupValid AND Initialized;
FEqualToleranceSubject.BindPublisher(Publisher := FCapture);
Initialized := FEqualToleranceSubject.Initialize(Parent := THIS^,
    AssertionName := 'EqualToleranceSubject');
FSetupValid := FSetupValid AND Initialized;
FNotEqualToleranceSubject.BindPublisher(Publisher := FCapture);
Initialized := FNotEqualToleranceSubject.Initialize(Parent := THIS^,
    AssertionName := 'NotEqualToleranceSubject');
FSetupValid := FSetupValid AND Initialized;
END_METHOD

{region 'Documentation'}
(*!
<summary>Establishes typed fixtures and verifies their representation before any subject call.</summary>
*)
{endregion}
METHOD PRIVATE InitializeValues : BOOL //! TRUE when fixture sizes and floating-point bit representations match their explicit expected patterns.
VAR
    Representation : FloatingPointBits_LReal;
END_VAR
Representation.Value := LREAL#1.0;
InitializeValues := (SIZEOF(Representation) = FixtureSize)
    AND (Representation.Bits = OneBits);

FQuietNaN.Bits := QuietNaNBits;
Representation.Value := FQuietNaN.Value;
InitializeValues := InitializeValues AND (Representation.Bits = QuietNaNBits);
FPositiveInfinity.Bits := PositiveInfinityBits;
Representation.Value := FPositiveInfinity.Value;
InitializeValues := InitializeValues AND (Representation.Bits = PositiveInfinityBits);
FNegativeInfinity.Bits := NegativeInfinityBits;
Representation.Value := FNegativeInfinity.Value;
InitializeValues := InitializeValues AND (Representation.Bits = NegativeInfinityBits);
END_METHOD

{region 'Documentation'}
(*!
<summary>Reads a captured finding; the caller bounds the index by 5 subjects.</summary>
*)
{endregion}
METHOD PRIVATE IsFindingValid : BOOL //! TRUE when the selected captured finding satisfies the scenario metadata and diagnostic checks.
VAR_INPUT
    Index : UINT; //! One-based index in the retained isolated event capture.
    ExpectedName : STRING(GVL_Constants.NameLength); //! Independently authored Assertion name expected in the selected finding.
    ExpectedResult : E_Result; //! Independently authored finding result.
END_VAR
IsFindingValid := (FEvents[Index].SequenceId = UINT_TO_UDINT(Index))
    AND (FEvents[Index].Name = ExpectedName)
    AND (FEvents[Index].OwnerScope = E_OwnerScope.Assertion)
    AND (FEvents[Index].EventType = E_EventType.Result)
    AND (FEvents[Index].State = E_State.Running)
    AND (FEvents[Index].Result = ExpectedResult)
    AND (FEvents[Index].Message <> '');
END_METHOD

{region 'Documentation'}
(*!
<summary>Completes abort without asynchronous resources.</summary>
*)
{endregion}
METHOD PROTECTED ProcessAbort
VAR_INPUT
    Enable : BOOL; //! Phase permission supplied by the owning Test Case; FALSE does not authorize progression, while observation may continue.
END_VAR
IF Enable THEN
    CompleteAbort();
END_IF;
END_METHOD

{region 'Documentation'}
(*!
<summary>Latches checked observations before the next script step may proceed.</summary>
*)
{endregion}
METHOD PROTECTED ProcessAssertions
VAR_INPUT
    Enable : BOOL; //! Phase permission supplied by the owning Test Case; FALSE does not authorize progression, while observation may continue.
END_VAR
VAR
    Evaluate : BOOL;
END_VAR
Evaluate := Enable AND FObservationReady;
FEqualResult(Enable := Evaluate,
    State := State,
    IN := FEqualResultMatches);
FLessThanResult(Enable := Evaluate,
    State := State,
    IN := FLessThanResultMatches);
FInRangeResult(Enable := Evaluate,
    State := State,
    IN := FInRangeResultMatches);
FEqualToleranceResult(Enable := Evaluate,
    State := State,
    IN := FEqualToleranceResultMatches);
FNotEqualToleranceResult(Enable := Evaluate,
    State := State,
    IN := FNotEqualToleranceResultMatches);
FCaptureIntegrity(Enable := Evaluate,
    State := State,
    IN := FCaptureIntegrityMatches);
FFindingDetails(Enable := Evaluate,
    State := State,
    IN := FFindingDetailsMatch);
IF Evaluate THEN
    FChecked := TRUE;
END_IF;
END_METHOD

{region 'Documentation'}
(*!
<summary>No Preparation phase is required.</summary>
*)
{endregion}
METHOD PROTECTED ProcessPreparations
VAR_INPUT
    // SA0033: Required hook; this test has no Preparation phase.
    {attribute 'analysis' := '-33'}
    Enable : BOOL; //! Phase permission supplied by the owning Test Case; FALSE does not authorize progression, while observation may continue.
END_VAR
END_METHOD

{region 'Documentation'}
(*!
<summary>Restarts the script and resets the checking Assertions.</summary>
*)
{endregion}
METHOD PROTECTED ProcessReset
FRow := ActualQuietNaN;
FRowPrepared := FALSE;
FChecked := FALSE;
FObservationReady := FALSE;
FEqualResult.Reset();
FEqualResultMatches := TRUE;
FLessThanResult.Reset();
FLessThanResultMatches := TRUE;
FInRangeResult.Reset();
FInRangeResultMatches := TRUE;
FEqualToleranceResult.Reset();
FEqualToleranceResultMatches := TRUE;
FNotEqualToleranceResult.Reset();
FNotEqualToleranceResultMatches := TRUE;
FCaptureIntegrity.Reset();
FCaptureIntegrityMatches := TRUE;
FFindingDetails.Reset();
FFindingDetailsMatch := TRUE;
CompleteReset();
END_METHOD

{region 'Documentation'}
(*!
<summary>Advances one bounded script step per active PLC cycle.</summary>
*)
{endregion}
METHOD PROTECTED ProcessTests
VAR_INPUT
    Enable : BOOL; //! Phase permission supplied by the owning Test Case; FALSE does not authorize progression, while observation may continue.
END_VAR
IF NOT Enable THEN
    RETURN;
END_IF;

IF FChecked THEN
    FChecked := FALSE;
    FObservationReady := FALSE;
    IF FRow = LastRow THEN
        CompleteTests();
        RETURN;
    END_IF;
    FRow := FRow + 1;
    FRowPrepared := FALSE;
END_IF;

IF NOT FRowPrepared THEN
    SelectRow();
    FCapture.Reset();
    IF NOT FPreserveResults THEN
        ResetSubjects();
    END_IF;
    CallSubjects(Enable := FALSE);
    FRowPrepared := TRUE;
ELSE
    CallSubjects(Enable := TRUE);
    CheckResults();
    FObservationReady := TRUE;
END_IF;
END_METHOD

{region 'Documentation'}
(*!
<summary>Requests fresh subject results before the next disabled call.</summary>
*)
{endregion}
METHOD PRIVATE ResetSubjects
FEqualSubject.Reset();
FLessThanSubject.Reset();
FInRangeSubject.Reset();
FEqualToleranceSubject.Reset();
FNotEqualToleranceSubject.Reset();
END_METHOD

